(* IEC 61131-3 sources: 2026_Projet_YGO_ExcavatriceDragage/TOOLS/TEST_AUTO_CI/RESULTS/G_CYCLE/reports (part 2) *)

(* ---- FB_CycleSemiAuto_test.st ---- *)
SETUP
VAR
    FB : FB_CycleSemiAuto;
    SampleCount : INT := 0;
    SampleCountTotal : UDINT := 0;
END_VAR
END_SETUP

TEST 'T262-002 AX10B : transfert Both P1 sans coupure M2 puis AX11 P2'
    (* Chargement securise de AX10B : consigne de forcage ecrite par l'operateur (T358). *)
    FB(Enable := TRUE, PowerContactorEngaged := TRUE, Mode := E_Mode.SEMI_AUTO,
       HeartbeatIhmOk := TRUE, M1_SpeedValid := TRUE, M2_SpeedValid := TRUE,
       M1_ContactorsReleased := TRUE, M2_ContactorsReleased := TRUE,
       M1_BrakeApplied := TRUE, M2_BrakeApplied := TRUE,
       M1_MeasuredSpeedMps := 0.0, M2_MeasuredSpeedMps := 0.0,
       JoystickDeflected := FALSE, DeadmanArmed := FALSE,
       CfgCommissioningEnable := TRUE, CfgCtrlAscentMaxStep := 2,
       CfgCtrlAscentDistanceM := 2.0, SampleCount := SampleCount, StepForceTgt := 22);
    ASSERT_TRUE(FB.ForceStepAccepted, 'AX10B forcee immediatement (T358)');
    ASSERT_TRUE(FB.StepForceTgtTaken, 'Consigne vue par le FB : PRG_03 l acquitte (T358)');

    (* Scans d acquittement puis d execution : aucun mouvement au chargement. *)
    FB(StepForceTgt := -1, SampleCount := SampleCount);
    FB(SampleCount := SampleCount);
    ASSERT_FALSE(FB.WinchM1Cmd.RunRequest OR FB.WinchM2Cmd.RunRequest,
                 'Chargement AX10B sans mouvement');

    (* Nouveau geste Y+ : M1 et M2 sont publies simultanement a P1. *)
    FB(StartCycle := FALSE, JoystickDeflected := TRUE, DeadmanArmed := TRUE,
       JoystickPull := TRUE, M2_SpeedStepApplied := 1,
       M1FinalAscentStartReady := TRUE, Benne_CloseReached := TRUE,
       Benne_IsClosed := TRUE, Benne_IsRoughlyClosed := TRUE,
       SampleCount := SampleCount);
    ASSERT_TRUE(FB.CycleStep = E_AutoCycleStep.AX10B_RACCORDEMENT_P1,
                'Scan transfert execute en AX10B');
    ASSERT_TRUE(FB.WinchM1Cmd.RunRequest AND FB.WinchM2Cmd.RunRequest,
                'AX10B publie Both sans trou de commande');
    ASSERT_TRUE((FB.WinchM1Cmd.StepTgt = 1) AND (FB.WinchM2Cmd.StepTgt = 1),
                'AX10B publie M1 P1 et M2 P1');
    ASSERT_TRUE(FB.WinchM1Cmd.ReqAscent AND FB.WinchM2Cmd.ReqAscent,
                'AX10B conserve le sens montee des deux treuils');

    (* Scan suivant : AX11 reprend avec le plafond commun configure P2. *)
    FB(SampleCount := SampleCount);
    ASSERT_TRUE(FB.CycleStep = E_AutoCycleStep.AX11_CTRL_ASCENT,
                'AX11 prend le relais apres transfert P1/P1');
    ASSERT_TRUE((FB.WinchM1Cmd.StepTgt = 2) AND (FB.WinchM2Cmd.StepTgt = 2),
                'AX11 applique le plafond commun P2');
END_TEST

(* ============================================================================
   T345-L2 - AX14->AX15A instantane, neutre obligatoire avant AX15B
   Contrat : TASK_CONTRACT_T345_L2_AX14_AX15A_INSTANTANEE.yaml
   ============================================================================ *)

TEST 'T345-L2-001 : arrivee AX14 neutre, puis nouveau push autorise AX15B'
    FB(Enable := TRUE, PowerContactorEngaged := TRUE, Mode := E_Mode.SEMI_AUTO,
       HeartbeatIhmOk := TRUE, M1_SpeedValid := TRUE, M2_SpeedValid := TRUE,
       M1_ContactorsReleased := TRUE, M2_ContactorsReleased := TRUE,
       M1_BrakeApplied := TRUE, M2_BrakeApplied := TRUE,
       HomedM1 := TRUE, HomedM2 := TRUE, InitPositionOk := TRUE, WinchesAtTopWindow := TRUE,
       Translation_At_Tremie := TRUE, Translation_Busy := FALSE,
       JoystickDeflected := FALSE, DeadmanArmed := TRUE,
       JoystickPush := FALSE, JoystickPull := FALSE, JoystickLeft := FALSE, JoystickRight := FALSE,
       SampleCount := SampleCount, StepForceTgt := 14);
    ASSERT_TRUE(FB.ForceStepAccepted, 'T345-L2-001 : AX14 force');
    FB(StepForceTgt := -1, Translation_At_Tremie := TRUE, Translation_Busy := FALSE,
       JoystickDeflected := FALSE, DeadmanArmed := TRUE, JoystickPush := FALSE,
       SampleCount := SampleCount);
    ADVANCE_TIME(600000000);
    FB(Translation_At_Tremie := TRUE, Translation_Busy := FALSE,
       JoystickDeflected := FALSE, DeadmanArmed := TRUE, JoystickPush := FALSE,
       SampleCount := SampleCount);

    (* Premier scan AX15A au neutre : le latch s'arme, sans transition dans ce meme scan. *)
    FB(Translation_At_Tremie := TRUE, Translation_Busy := FALSE,
       JoystickDeflected := FALSE, DeadmanArmed := TRUE, JoystickPush := FALSE,
       SampleCount := SampleCount);
    ASSERT_TRUE(FB.CycleStep = E_AutoCycleStep.AX15A_DUMP_ARRIVE,
                'T345-L2-001 : AX15A atteint apres confirmation arret');
    ASSERT_FALSE(FB.BucketCmd.ReqOpen OR FB.WinchM1Cmd.RunRequest OR FB.WinchM2Cmd.RunRequest OR FB.TranslationCmd.ReqStart,
                 'T345-L2-001 : aucune commande au scan neutre AX15A');
    ASSERT_EQ(FB.OperatorAction, 'AX15a - Pousser vers le bas pour ouvrir et vider.',
              'T345-L2-001 : guide push publie apres neutre');

    (* Nouveau geste : changement d'etat, puis commande seulement au scan AX15B. *)
    FB(JoystickDeflected := TRUE, DeadmanArmed := TRUE, JoystickPush := TRUE,
       SampleCount := SampleCount);
    ASSERT_TRUE(FB.CycleStep = E_AutoCycleStep.AX15A_DUMP_ARRIVE,
                'T345-L2-001 : transition demandee depuis AX15A');
    ASSERT_FALSE(FB.BucketCmd.ReqOpen, 'T345-L2-001 : aucune ouverture au scan de transition');
    FB(JoystickDeflected := TRUE, DeadmanArmed := TRUE, JoystickPush := TRUE,
       SampleCount := SampleCount);
    ASSERT_TRUE(FB.CycleStep = E_AutoCycleStep.AX15B_DUMP_OPEN,
                'T345-L2-001 : AX15B execute au scan suivant');
    ASSERT_TRUE(FB.BucketCmd.ReqOpen, 'T345-L2-001 : ouverture autorisee apres neutre puis nouveau push');
END_TEST

TEST 'T345-L2-002 : push Y maintenu a l arrivee passe AX15A mais reste bloque avant neutre'
    FB(Enable := TRUE, PowerContactorEngaged := TRUE, Mode := E_Mode.SEMI_AUTO,
       HeartbeatIhmOk := TRUE, M1_SpeedValid := TRUE, M2_SpeedValid := TRUE,
       M1_ContactorsReleased := TRUE, M2_ContactorsReleased := TRUE,
       M1_BrakeApplied := TRUE, M2_BrakeApplied := TRUE,
       HomedM1 := TRUE, HomedM2 := TRUE, InitPositionOk := TRUE, WinchesAtTopWindow := TRUE,
       Translation_At_Tremie := TRUE, Translation_Busy := FALSE,
       JoystickDeflected := TRUE, DeadmanArmed := TRUE,
       JoystickPush := TRUE, JoystickPull := FALSE, JoystickLeft := FALSE, JoystickRight := FALSE,
       SampleCount := SampleCount, StepForceTgt := 14);
    FB(StepForceTgt := -1, Translation_At_Tremie := TRUE, Translation_Busy := FALSE,
       JoystickDeflected := TRUE, DeadmanArmed := TRUE, JoystickPush := TRUE,
       SampleCount := SampleCount);
    ADVANCE_TIME(600000000);
    FB(Translation_At_Tremie := TRUE, Translation_Busy := FALSE,
       JoystickDeflected := TRUE, DeadmanArmed := TRUE, JoystickPush := TRUE,
       SampleCount := SampleCount);
    FB(Translation_At_Tremie := TRUE, Translation_Busy := FALSE,
       JoystickDeflected := TRUE, DeadmanArmed := TRUE, JoystickPush := TRUE,
       SampleCount := SampleCount);
    ASSERT_TRUE(FB.CycleStep = E_AutoCycleStep.AX15A_DUMP_ARRIVE,
                'T345-L2-002 : transition AX14->AX15A sans attendre neutre');
    ASSERT_TRUE(FB.WaitingForOperator, 'T345-L2-002 : relachement operateur attendu');
    ASSERT_EQ(FB.OperatorAction, 'AX15a - Relacher le joystick avant ouverture.',
              'T345-L2-002 : message de relachement explicite');
    ASSERT_FALSE(FB.BucketCmd.ReqOpen OR FB.WinchM1Cmd.RunRequest OR FB.WinchM2Cmd.RunRequest OR FB.TranslationCmd.ReqStart,
                 'T345-L2-002 : Y maintenu ne commande aucun mouvement avant neutre');
    FB(JoystickDeflected := TRUE, DeadmanArmed := TRUE, JoystickPush := TRUE,
       SampleCount := SampleCount);
    ASSERT_TRUE(FB.CycleStep = E_AutoCycleStep.AX15A_DUMP_ARRIVE,
                'T345-L2-002 : AX15A maintenu tant que Y reste pousse');
    ASSERT_FALSE(FB.BucketCmd.ReqOpen, 'T345-L2-002 : ReqOpen reste faux avant neutre');
END_TEST

TEST 'T345-L2-003 : diagonale X plus Y maintenue ne contourne pas le neutre AX15A'
    FB(Enable := TRUE, PowerContactorEngaged := TRUE, Mode := E_Mode.SEMI_AUTO,
       HeartbeatIhmOk := TRUE, M1_SpeedValid := TRUE, M2_SpeedValid := TRUE,
       M1_ContactorsReleased := TRUE, M2_ContactorsReleased := TRUE,
       M1_BrakeApplied := TRUE, M2_BrakeApplied := TRUE,
       HomedM1 := TRUE, HomedM2 := TRUE, InitPositionOk := TRUE, WinchesAtTopWindow := TRUE,
       Translation_At_Tremie := TRUE, Translation_Busy := FALSE,
       JoystickDeflected := TRUE, DeadmanArmed := TRUE,
       JoystickPush := TRUE, JoystickPull := FALSE, JoystickLeft := TRUE, JoystickRight := FALSE,
       SampleCount := SampleCount, StepForceTgt := 14);
    FB(StepForceTgt := -1, Translation_At_Tremie := TRUE, Translation_Busy := FALSE,
       JoystickDeflected := TRUE, DeadmanArmed := TRUE, JoystickPush := TRUE, JoystickLeft := TRUE,
       SampleCount := SampleCount);
    ADVANCE_TIME(600000000);
    FB(Translation_At_Tremie := TRUE, Translation_Busy := FALSE,
       JoystickDeflected := TRUE, DeadmanArmed := TRUE, JoystickPush := TRUE, JoystickLeft := TRUE,
       SampleCount := SampleCount);
    FB(Translation_At_Tremie := TRUE, Translation_Busy := FALSE,
       JoystickDeflected := TRUE, DeadmanArmed := TRUE, JoystickPush := TRUE, JoystickLeft := TRUE,
       SampleCount := SampleCount);
    ASSERT_TRUE(FB.CycleStep = E_AutoCycleStep.AX15A_DUMP_ARRIVE,
                'T345-L2-003 : diagonale n empeche pas l arrivee AX15A');
    ASSERT_FALSE(FB.BucketCmd.ReqOpen OR FB.WinchM1Cmd.RunRequest OR FB.WinchM2Cmd.RunRequest OR FB.TranslationCmd.ReqStart,
                 'T345-L2-003 : diagonale ne produit aucun mouvement avant neutre');
    FB(JoystickDeflected := TRUE, DeadmanArmed := TRUE, JoystickPush := TRUE, JoystickLeft := TRUE,
       SampleCount := SampleCount);
    ASSERT_TRUE(FB.CycleStep = E_AutoCycleStep.AX15A_DUMP_ARRIVE,
                'T345-L2-003 : diagonale maintenue reste bloquee en AX15A');
    ASSERT_FALSE(FB.BucketCmd.ReqOpen, 'T345-L2-003 : ReqOpen reste faux sous diagonale');
END_TEST

TEST 'T345-L2-004 : forcage repete cible 15 efface un latch neutre precedent'
    FB(Enable := TRUE, PowerContactorEngaged := TRUE, Mode := E_Mode.SEMI_AUTO,
       HeartbeatIhmOk := TRUE, M1_SpeedValid := TRUE, M2_SpeedValid := TRUE,
       M1_ContactorsReleased := TRUE, M2_ContactorsReleased := TRUE,
       M1_BrakeApplied := TRUE, M2_BrakeApplied := TRUE,
       HomedM1 := TRUE, HomedM2 := TRUE, InitPositionOk := TRUE, WinchesAtTopWindow := TRUE,
       JoystickDeflected := FALSE, DeadmanArmed := TRUE, JoystickPush := FALSE,
       SampleCount := SampleCount, StepForceTgt := 15);
    FB(StepForceTgt := -1, JoystickDeflected := FALSE, DeadmanArmed := TRUE, JoystickPush := FALSE,
       SampleCount := SampleCount);
    ASSERT_TRUE(FB.CycleStep = E_AutoCycleStep.AX15A_DUMP_ARRIVE,
                'T345-L2-004 : AX15A execute au neutre et latch arme');

    (* Meme cible forcee pendant un push : le reset doit avoir lieu meme sans changement d enum. *)
    FB(StepForceTgt := 15, JoystickDeflected := TRUE, DeadmanArmed := TRUE, JoystickPush := TRUE,
       SampleCount := SampleCount);
    ASSERT_TRUE(FB.ForceStepAccepted, 'T345-L2-004 : forcage repete 15 accepte et neutre en commandes');
    ASSERT_FALSE(FB.BucketCmd.ReqOpen, 'T345-L2-004 : scan de forcage sans ouverture');
    FB(StepForceTgt := -1, JoystickDeflected := TRUE, DeadmanArmed := TRUE, JoystickPush := TRUE,
       SampleCount := SampleCount);
    FB(JoystickDeflected := TRUE, DeadmanArmed := TRUE, JoystickPush := TRUE,
       SampleCount := SampleCount);
    ASSERT_TRUE(FB.CycleStep = E_AutoCycleStep.AX15A_DUMP_ARRIVE,
                'T345-L2-004 : latch perime ne survit pas au forcage repete');
    ASSERT_FALSE(FB.BucketCmd.ReqOpen, 'T345-L2-004 : push deja actif reste bloque sans nouveau neutre');
END_TEST

TEST 'T345-L2-005 : non regression AX2 vers AX3 conserve le geste PushOnly existant'
    FB(Enable := TRUE, PowerContactorEngaged := TRUE, Mode := E_Mode.SEMI_AUTO,
       HeartbeatIhmOk := TRUE, M1_SpeedValid := TRUE, M2_SpeedValid := TRUE,
       M1_ContactorsReleased := TRUE, M2_ContactorsReleased := TRUE,
       M1_BrakeApplied := TRUE, M2_BrakeApplied := TRUE,
       HomedM1 := TRUE, HomedM2 := TRUE, InitPositionOk := TRUE, WinchesAtTopWindow := TRUE,
       Translation_At_P1 := TRUE, Translation_Busy := FALSE,
       JoystickDeflected := TRUE, DeadmanArmed := TRUE,
       JoystickPush := TRUE, JoystickPull := FALSE, JoystickLeft := FALSE, JoystickRight := FALSE,
       SampleCount := SampleCount, StepForceTgt := 2);
    FB(StepForceTgt := -1, Translation_At_P1 := TRUE, Translation_Busy := FALSE,
       JoystickDeflected := TRUE, DeadmanArmed := TRUE, JoystickPush := TRUE,
       JoystickLeft := FALSE, JoystickRight := FALSE, SampleCount := SampleCount);
    ADVANCE_TIME(600000000);
    FB(Translation_At_P1 := TRUE, Translation_Busy := FALSE,
       JoystickDeflected := TRUE, DeadmanArmed := TRUE, JoystickPush := TRUE,
       JoystickLeft := FALSE, JoystickRight := FALSE, SampleCount := SampleCount);
    FB(Translation_At_P1 := TRUE, Translation_Busy := FALSE,
       JoystickDeflected := TRUE, DeadmanArmed := TRUE, JoystickPush := TRUE,
       JoystickLeft := FALSE, JoystickRight := FALSE, SampleCount := SampleCount);
    ASSERT_TRUE(FB.CycleStep = E_AutoCycleStep.AX3_OPEN_BUCKET,
                'T345-L2-005 : AX2->AX3 PushOnly inchange');
    ASSERT_TRUE(FB.BucketCmd.ReqOpen, 'T345-L2-005 : AX3 ouvre comme avant');
END_TEST

TEST 'T262-003 AX10B : timeout M1 borne a 2 s puis repli sans redemarrage implicite'
    (* Preparation AX10B au neutre, comme pour le test nominal (T358). *)
    FB(Enable := TRUE, PowerContactorEngaged := TRUE, Mode := E_Mode.SEMI_AUTO,
       HeartbeatIhmOk := TRUE, M1_SpeedValid := TRUE, M2_SpeedValid := TRUE,
       M1_ContactorsReleased := TRUE, M2_ContactorsReleased := TRUE,
       M1_BrakeApplied := TRUE, M2_BrakeApplied := TRUE,
       M1_MeasuredSpeedMps := 0.0, M2_MeasuredSpeedMps := 0.0,
       JoystickDeflected := FALSE, DeadmanArmed := FALSE,
       CfgCommissioningEnable := TRUE, CfgCtrlAscentMaxStep := 2,
       CfgCtrlAscentDistanceM := 2.0, SampleCount := SampleCount, StepForceTgt := 22);
    ASSERT_TRUE(FB.ForceStepAccepted, 'AX10B forcee pour test timeout (T358)');
    ASSERT_TRUE(FB.StepForceTgtTaken, 'Consigne vue par le FB : PRG_03 l acquitte (T358)');
    FB(StepForceTgt := -1, SampleCount := SampleCount);
    FB(SampleCount := SampleCount);

    (* M1 indisponible : M2 est tenu en P1 pendant la fenetre bornee. *)
    FB(StartCycle := FALSE, JoystickDeflected := TRUE, DeadmanArmed := TRUE,
       JoystickPull := TRUE, M2_SpeedStepApplied := 1,
       M1FinalAscentStartReady := FALSE, Benne_CloseReached := TRUE,
       Benne_IsClosed := TRUE, Benne_IsRoughlyClosed := TRUE,
       SampleCount := SampleCount);
    ASSERT_TRUE(FB.BucketCmd.ReqHoldAscentP1AfterClose,
                'Fenetre AX10B : maintien P1 actif avant timeout');

    ADVANCE_TIME(2100000000);
    FB(SampleCount := SampleCount);
    ASSERT_FALSE(FB.BucketCmd.ReqHoldAscentP1AfterClose,
                 'Timeout : maintien M2 libere');
    ASSERT_FALSE(FB.WinchM1Cmd.RunRequest OR FB.WinchM2Cmd.RunRequest,
                 'Timeout : aucun redemarrage pendant arret de repli');

    ADVANCE_TIME(600000000);
    FB(SampleCount := SampleCount);
    ASSERT_TRUE(FB.CycleStep = E_AutoCycleStep.AX10B_RACCORDEMENT_P1,
                'Repli : AX10B conserve la main pendant la confirmation arret');
    ADVANCE_TIME(600000000);
    FB(SampleCount := SampleCount);
    ASSERT_TRUE(FB.CycleStep = E_AutoCycleStep.AX10B_RACCORDEMENT_P1,
                'Repli : dernier scan AX10B avant reprise');
    FB(SampleCount := SampleCount);
    ASSERT_TRUE(FB.CycleStep = E_AutoCycleStep.AX11_CTRL_ASCENT,
                'Repli : reprise explicite par AX11');
    ASSERT_TRUE(FB.WinchM1Cmd.RunRequest AND FB.WinchM2Cmd.RunRequest,
                'Repli : AX11 reprend les deux treuils ensemble');
END_TEST

TEST 'T331-001 AX15d micro-step benne : tirer ouvre le module, pousser ouvrir, relacher retour AX15B'
    SampleCount := 0;

    (* Chargement securise de l etape de vidage au joystick neutre, machine arretee. *)
    FB(Enable := TRUE, Reset := FALSE, PowerContactorEngaged := TRUE, Mode := E_Mode.SEMI_AUTO,
       HeartbeatIhmOk := TRUE, M1_SpeedValid := TRUE, M2_SpeedValid := TRUE,
       M1_ContactorsReleased := TRUE, M2_ContactorsReleased := TRUE,
       M1_BrakeApplied := TRUE, M2_BrakeApplied := TRUE,
       M1_MeasuredSpeedMps := 0.0, M2_MeasuredSpeedMps := 0.0,
       M1_SpeedStepApplied := 1, M2_SpeedStepApplied := 1,
       JoystickDeflected := FALSE, DeadmanArmed := FALSE,
       JoystickPush := FALSE, JoystickPull := FALSE, JoystickRight := FALSE, JoystickLeft := FALSE,
       StartCycle := FALSE, AbortCycle := FALSE,
       SpeedMismatchThresholdMps := 0.0, SpeedMismatchTimeout := T#0ms,
       WinchSyncError := FALSE, WinchSyncDeltaM := 0.0,
       HomedM1 := TRUE, HomedM2 := TRUE, InitPositionOk := TRUE, WinchesAtTopWindow := TRUE,
       M1_CablePosM := 7.0, M2_CablePosM := 7.0,
       Translation_At_P1 := FALSE, Translation_At_Tremie := TRUE, Translation_At_Maintenance := FALSE,
       Translation_Busy := FALSE, Translation_Done := TRUE,
       Benne_Busy := FALSE, Benne_Done := FALSE, Benne_CloseReached := FALSE,
       Benne_IsOpen := FALSE, Benne_IsClosed := FALSE, Benne_IsRoughlyClosed := FALSE,
       RepositionRequest := FALSE, SkipDrainRequest := FALSE, CfgDrainTime := T#0s,
       CfgCommissioningEnable := TRUE,
       CfgCtrlAscentMaxStep := 1, CfgCtrlAscentDistanceM := 2.0,
       SampleCount := SampleCount);
    FB(StepForceTgt := 16, SampleCount := SampleCount);
    ASSERT_TRUE(FB.ForceStepAccepted, 'Etape de vidage forcee (T331-001)');
    FB(StepForceTgt := -1, SampleCount := SampleCount);
    FB(SampleCount := SampleCount);

    (* Geste nominal maintenu Y- : vidage, treuils neutralises, aucune transition. *)
    FB(StartCycle := FALSE, JoystickDeflected := TRUE, DeadmanArmed := TRUE,
       JoystickPush := TRUE, SampleCount := SampleCount);
    ASSERT_TRUE(FB.CycleStep = E_AutoCycleStep.AX15B_DUMP_OPEN, 'Vidage observe');
    ASSERT_TRUE(FB.BucketCmd.ReqOpen, 'Vidage : ouverture benne commandee');
    ASSERT_FALSE(FB.BucketCmd.ReqClose, 'Vidage : aucune fermeture benne commandee');
    ASSERT_FALSE(FB.WinchM1Cmd.RunRequest OR FB.WinchM2Cmd.RunRequest,
                 'Vidage : les deux treuils restent neutralises');

    (* T383 : tirer ne fait PLUS de saut AX15B -> AX10. Il entre dans le micro-step AX15D. *)
    FB(JoystickPush := FALSE, JoystickPull := TRUE, SampleCount := SampleCount);
    FB(SampleCount := SampleCount);
    ASSERT_TRUE(FB.CycleStep = E_AutoCycleStep.AX15D_DUMP_BUCKET_JOG,
                'T383 : tirer entre dans le micro-step benne AX15D');
    ASSERT_FALSE(FB.CycleStep = E_AutoCycleStep.AX10_CLOSE_BUCKET,
                 'T383 : AUCUN saut vers AX10 (decharge non declaree retiree)');
    ASSERT_FALSE(FB.BucketCmd.ReqOpen, 'AX15D : ouverture neutralisee au tirer');
    ASSERT_TRUE(FB.BucketCmd.ReqClose, 'AX15D : tirer ferme la benne');
    ASSERT_FALSE(FB.WinchM1Cmd.RunRequest OR FB.WinchM2Cmd.RunRequest,
                 'AX15D : les deux treuils restent a 0 (aucun mouvement)');

    (* Module : pousser dans AX15D rouvre la benne, treuils toujours 0. *)
    FB(JoystickPush := TRUE, JoystickPull := FALSE, SampleCount := SampleCount);
    ASSERT_TRUE(FB.CycleStep = E_AutoCycleStep.AX15D_DUMP_BUCKET_JOG,
                'AX15D : on reste dans le micro-step pendant la manipulation');
    ASSERT_TRUE(FB.BucketCmd.ReqOpen, 'AX15D : pousser ouvre la benne');
    ASSERT_FALSE(FB.BucketCmd.ReqClose, 'AX15D : aucune fermeture simultanee');
    ASSERT_FALSE(FB.WinchM1Cmd.RunRequest OR FB.WinchM2Cmd.RunRequest,
                 'AX15D : treuils neutralises pendant le module');

    (* Retour au centre mort : on reprend le vidage (AX15B) sans remontee. *)
    FB(JoystickPush := FALSE, JoystickPull := FALSE, JoystickDeflected := FALSE,
       SampleCount := SampleCount);
    FB(SampleCount := SampleCount);   // AX15D assigne State:=AX15B -> CycleStep au scan suivant
    ASSERT_TRUE(FB.CycleStep = E_AutoCycleStep.AX15B_DUMP_OPEN,
                'AX15D : relachement -> retour au vidage AX15B');
    ASSERT_FALSE(FB.BucketCmd.ReqOpen OR FB.BucketCmd.ReqClose,
                 'AX15D : neutre = les deux demandes benne a zero');
    ASSERT_FALSE(FB.WinchM1Cmd.RunRequest OR FB.WinchM2Cmd.RunRequest,
                 'AX15D : aucun treuil commande au relachement');

    (* Fin de vidage : la benne ouverte amene AX18 sur geste pousse, inchange. *)
    FB(Benne_Done := TRUE, Benne_IsOpen := TRUE, Benne_IsClosed := FALSE,
       Benne_IsRoughlyClosed := FALSE, JoystickDeflected := TRUE, JoystickPush := TRUE,
       SampleCount := SampleCount);
    FB(SampleCount := SampleCount);
    ASSERT_TRUE(FB.CycleStep = E_AutoCycleStep.AX18_DONE_SYNC,
                'Fin de vidage apres module : AX18 inchange');
    ASSERT_FALSE(FB.BucketCmd.ReqOpen, 'Fin de vidage : ouverture relachee');
END_TEST

TEST 'T331-002 AX15b/AX15c non-regression : vidage nominal et repositionnement inchanges'
    SampleCount := 0;

    (* Chargement securise de l etape de vidage au joystick neutre. *)
    FB(Enable := TRUE, Reset := FALSE, PowerContactorEngaged := TRUE, Mode := E_Mode.SEMI_AUTO,
       HeartbeatIhmOk := TRUE, M1_SpeedValid := TRUE, M2_SpeedValid := TRUE,
       M1_ContactorsReleased := TRUE, M2_ContactorsReleased := TRUE,
       M1_BrakeApplied := TRUE, M2_BrakeApplied := TRUE,
       M1_MeasuredSpeedMps := 0.0, M2_MeasuredSpeedMps := 0.0,
       M1_SpeedStepApplied := 1, M2_SpeedStepApplied := 1,
       JoystickDeflected := FALSE, DeadmanArmed := FALSE,
       JoystickPush := FALSE, JoystickPull := FALSE, JoystickRight := FALSE, JoystickLeft := FALSE,
       StartCycle := FALSE, AbortCycle := FALSE,
       SpeedMismatchThresholdMps := 0.0, SpeedMismatchTimeout := T#0ms,
       WinchSyncError := FALSE, WinchSyncDeltaM := 0.0,
       HomedM1 := TRUE, HomedM2 := TRUE, InitPositionOk := TRUE, WinchesAtTopWindow := TRUE,
       M1_CablePosM := 7.0, M2_CablePosM := 7.0,
       Translation_At_P1 := FALSE, Translation_At_Tremie := TRUE, Translation_At_Maintenance := FALSE,
       Translation_Busy := FALSE, Translation_Done := TRUE,
       Benne_Busy := FALSE, Benne_Done := FALSE, Benne_CloseReached := FALSE,
       Benne_IsOpen := FALSE, Benne_IsClosed := FALSE, Benne_IsRoughlyClosed := FALSE,
       RepositionRequest := FALSE, SkipDrainRequest := FALSE, CfgDrainTime := T#0s,
       CfgCommissioningEnable := TRUE,
       CfgCtrlAscentMaxStep := 1, CfgCtrlAscentDistanceM := 2.0,
       SampleCount := SampleCount);
    FB(StepForceTgt := 16, SampleCount := SampleCount);
    ASSERT_TRUE(FB.ForceStepAccepted, 'Etape de vidage forcee (non-regression T358)');
    ASSERT_TRUE(FB.StepForceTgtTaken, 'Consigne vue par le FB : PRG_03 l acquitte (T358)');
    FB(StepForceTgt := -1, SampleCount := SampleCount);

    (* Vidage nominal Y- : ouverture seule, treuils neutralises. *)
    FB(StartCycle := FALSE, JoystickDeflected := TRUE, DeadmanArmed := TRUE,
       JoystickPush := TRUE, SampleCount := SampleCount);
    ASSERT_TRUE(FB.CycleStep = E_AutoCycleStep.AX15B_DUMP_OPEN, 'Vidage nominal inchange');
    ASSERT_TRUE(FB.BucketCmd.ReqOpen, 'Vidage nominal : ouverture commandee');
    ASSERT_FALSE(FB.BucketCmd.ReqClose, 'Vidage nominal : aucune fermeture');
    ASSERT_FALSE(FB.WinchM1Cmd.RunRequest OR FB.WinchM2Cmd.RunRequest,
                 'Vidage nominal : treuils a l arret');

    (* Option IHM maintenue : repositionnement couple en descente, inchange. *)
    FB(RepositionRequest := TRUE, SampleCount := SampleCount);
    FB(SampleCount := SampleCount);
    ASSERT_TRUE(FB.CycleStep = E_AutoCycleStep.AX15C_DUMP_REPOSITION,
                'Repositionnement inchange : AX15c atteint');
    ASSERT_TRUE(FB.WinchM1Cmd.RunRequest AND FB.WinchM2Cmd.RunRequest,
                'Repositionnement : M1 et M2 commandes');
    ASSERT_TRUE(FB.WinchM1Cmd.ReqDescend AND FB.WinchM2Cmd.ReqDescend,
                'Repositionnement : descente couplee conservee');
    ASSERT_FALSE(FB.WinchM1Cmd.ReqAscent OR FB.WinchM2Cmd.ReqAscent,
                 'Repositionnement : aucune montee commandee');
    ASSERT_EQ(FB.WinchM1Cmd.StepTgt, FB.WinchM2Cmd.StepTgt,
              'Repositionnement : meme palier M1/M2');

    (* Relachement de l option : retour au vidage, treuils de nouveau a l arret. *)
    FB(RepositionRequest := FALSE, SampleCount := SampleCount);
    FB(SampleCount := SampleCount);
    ASSERT_TRUE(FB.CycleStep = E_AutoCycleStep.AX15B_DUMP_OPEN,
                'Retour au vidage inchange au relachement de l option');
    ASSERT_FALSE(FB.WinchM1Cmd.RunRequest OR FB.WinchM2Cmd.RunRequest,
                 'Retour vidage : treuils arretes');

    (* Vidage termine : la benne ouverte amene la fin de passe, inchange. *)
    FB(Benne_Done := TRUE, Benne_IsOpen := TRUE, Benne_IsClosed := FALSE,
       Benne_IsRoughlyClosed := FALSE, SampleCount := SampleCount);
    FB(SampleCount := SampleCount);
    ASSERT_TRUE(FB.CycleStep = E_AutoCycleStep.AX18_DONE_SYNC, 'Fin de vidage inchangee');
    ASSERT_FALSE(FB.BucketCmd.ReqOpen, 'Fin de vidage : ouverture relachee');
    ASSERT_EQ(FB.SampleCount, 1, 'Fin de vidage : compteur incremente une seule fois');
END_TEST

TEST 'T331-003 AX15d micro-step : perte du geste, de l homme-mort ou defaut neutralise sans reprise'
    SampleCount := 0;

    (* Chargement securise de l etape de vidage au joystick neutre. *)
    FB(Enable := TRUE, Reset := FALSE, PowerContactorEngaged := TRUE, Mode := E_Mode.SEMI_AUTO,
       HeartbeatIhmOk := TRUE, M1_SpeedValid := TRUE, M2_SpeedValid := TRUE,
       M1_ContactorsReleased := TRUE, M2_ContactorsReleased := TRUE,
       M1_BrakeApplied := TRUE, M2_BrakeApplied := TRUE,
       M1_MeasuredSpeedMps := 0.0, M2_MeasuredSpeedMps := 0.0,
       M1_SpeedStepApplied := 1, M2_SpeedStepApplied := 1,
       JoystickDeflected := FALSE, DeadmanArmed := FALSE,
       JoystickPush := FALSE, JoystickPull := FALSE, JoystickRight := FALSE, JoystickLeft := FALSE,
       StartCycle := FALSE, AbortCycle := FALSE,
       SpeedMismatchThresholdMps := 0.0, SpeedMismatchTimeout := T#0ms,
       WinchSyncError := FALSE, WinchSyncDeltaM := 0.0,
       HomedM1 := TRUE, HomedM2 := TRUE, InitPositionOk := TRUE, WinchesAtTopWindow := TRUE,
       M1_CablePosM := 7.0, M2_CablePosM := 7.0,
       Translation_At_P1 := FALSE, Translation_At_Tremie := TRUE, Translation_At_Maintenance := FALSE,
       Translation_Busy := FALSE, Translation_Done := TRUE,
       Benne_Busy := FALSE, Benne_Done := FALSE, Benne_CloseReached := FALSE,
       Benne_IsOpen := FALSE, Benne_IsClosed := FALSE, Benne_IsRoughlyClosed := FALSE,
       RepositionRequest := FALSE, SkipDrainRequest := FALSE, CfgDrainTime := T#0s,
       CfgCommissioningEnable := TRUE,
       CfgCtrlAscentMaxStep := 1, CfgCtrlAscentDistanceM := 2.0,
       SampleCount := SampleCount);
    FB(StepForceTgt := 16, SampleCount := SampleCount);
    ASSERT_TRUE(FB.ForceStepAccepted, 'Etape de vidage forcee (T331-003)');
    FB(StepForceTgt := -1, SampleCount := SampleCount);
    FB(SampleCount := SampleCount);

    (* Vidage puis tirer maintenu : entre dans le micro-step AX15D, fermeture commandee. *)
    FB(StartCycle := FALSE, JoystickDeflected := TRUE, DeadmanArmed := TRUE,
       JoystickPush := TRUE, SampleCount := SampleCount);
    FB(JoystickPush := FALSE, JoystickPull := TRUE, SampleCount := SampleCount);
    FB(SampleCount := SampleCount);
    ASSERT_TRUE(FB.CycleStep = E_AutoCycleStep.AX15D_DUMP_BUCKET_JOG,
                'Micro-step : entree dans AX15D au tirer');
    ASSERT_TRUE(FB.BucketCmd.ReqClose, 'Micro-step : fermeture benne commandee au tirer');

    (* Relachement du manche : plus aucune demande, retour au vidage AX15B. *)
    FB(JoystickDeflected := FALSE, JoystickPull := FALSE, DeadmanArmed := TRUE,
       SampleCount := SampleCount);
    ASSERT_FALSE(FB.BucketCmd.ReqClose, 'Relachement : fermeture benne neutralisee');
    ASSERT_FALSE(FB.WinchM1Cmd.RunRequest OR FB.WinchM2Cmd.RunRequest,
                 'Relachement : treuils neutralises');
    FB(SampleCount := SampleCount);
    ASSERT_TRUE(FB.CycleStep = E_AutoCycleStep.AX15B_DUMP_OPEN,
                'Relachement : retour a AX15B (reprendre le vidage)');
    ASSERT_FALSE(FB.BucketCmd.ReqClose, 'Relachement : aucune reprise automatique');

    (* Geste repris (tirer) : retour dans le micro-step sous commande maintenue. *)
    FB(JoystickDeflected := TRUE, JoystickPull := TRUE, SampleCount := SampleCount);
    FB(SampleCount := SampleCount);
    ASSERT_TRUE(FB.CycleStep = E_AutoCycleStep.AX15D_DUMP_BUCKET_JOG,
                'Geste repris : retour dans AX15D');
    ASSERT_TRUE(FB.BucketCmd.ReqClose, 'Geste repris : fermeture benne reprise');

    (* Perte de l homme-mort : neutralisation complete, etape conservee. *)
    FB(DeadmanArmed := FALSE, SampleCount := SampleCount);
    ASSERT_FALSE(FB.BucketCmd.ReqClose OR FB.BucketCmd.ReqOpen
                 OR FB.WinchM1Cmd.RunRequest OR FB.WinchM2Cmd.RunRequest,
                 'Homme-mort perdu : plus aucune demande de mouvement');
    FB(SampleCount := SampleCount);
    ASSERT_TRUE(FB.CycleStep = E_AutoCycleStep.AX15D_DUMP_BUCKET_JOG,
                'Homme-mort perdu : etape conservee, aucune reprise automatique');

    (* Defaut pendant le micro-step : repli AX_STAB, sorties neutralisees. *)
    FB(DeadmanArmed := TRUE, HeartbeatIhmOk := FALSE, SampleCount := SampleCount);
    ASSERT_TRUE(FB.CycleStep = E_AutoCycleStep.AX_STAB, 'Defaut : repli AX_STAB');
    ASSERT_FALSE(FB.BucketCmd.ReqClose OR FB.BucketCmd.ReqOpen
                 OR FB.WinchM1Cmd.RunRequest OR FB.WinchM2Cmd.RunRequest,
                 'Defaut : toutes les demandes neutralisees');
    ASSERT_FALSE(FB.Lifecycle.Busy, 'Defaut : cycle non actif');

    (* Acquittement conscient : cause disparue puis Reset. *)
    FB(HeartbeatIhmOk := TRUE, JoystickDeflected := FALSE, JoystickPull := FALSE,
       DeadmanArmed := FALSE, Reset := TRUE, SampleCount := SampleCount);
    FB(Reset := FALSE, SampleCount := SampleCount);
    ASSERT_FALSE(FB.Fault.Latched, 'Acquittement : defaut efface apres cause disparue');
    ASSERT_TRUE(FB.CycleStep = E_AutoCycleStep.AX0_REPOS, 'Acquittement : retour au repos');
END_TEST

TEST 'TC-P03-001 Dynamique Enable : neutralisation initiale, transition Ready au repos, puis coupure'
    (* Scan 0 : Enable=FALSE -> Neutralisation *)
    FB(Enable := FALSE, Reset := FALSE, PowerContactorEngaged := TRUE, Mode := E_Mode.SEMI_AUTO,
       DeadmanArmed := FALSE, JoystickDeflected := FALSE, JoystickPush := FALSE, M1_SpeedValid := TRUE, M2_SpeedValid := TRUE, M1_ContactorsReleased := TRUE, M2_ContactorsReleased := TRUE, M1_BrakeApplied := TRUE, M2_BrakeApplied := TRUE, M1_SpeedStepApplied := 4, M2_SpeedStepApplied := 4, HeartbeatIhmOk := TRUE,
       StartCycle := FALSE, SampleCount := SampleCount);
    ASSERT_FALSE(FB.Ready, 'Enable=FALSE -> Ready=FALSE (neutralise)');
    ASSERT_FALSE(FB.Lifecycle.Busy, 'Enable=FALSE -> Lifecycle.Busy=FALSE');

    ADVANCE_TIME(10000000);

    (* Scan 1 : Enable=TRUE -> Prete en service *)
    FB(Enable := TRUE, Reset := FALSE, PowerContactorEngaged := TRUE, Mode := E_Mode.SEMI_AUTO,
       DeadmanArmed := FALSE, JoystickDeflected := FALSE, JoystickPush := FALSE, M1_SpeedValid := TRUE, M2_SpeedValid := TRUE, M1_ContactorsReleased := TRUE, M2_ContactorsReleased := TRUE, M1_BrakeApplied := TRUE, M2_BrakeApplied := TRUE, M1_SpeedStepApplied := 4, M2_SpeedStepApplied := 4, HeartbeatIhmOk := TRUE,
       StartCycle := FALSE, SampleCount := SampleCount);
    ASSERT_TRUE(FB.Ready, 'Enable=TRUE -> Ready=TRUE (nominal)');
    ASSERT_FALSE(FB.Lifecycle.Busy, 'Au repos -> Pas de cycle actif');

    ADVANCE_TIME(10000000);

    (* Scan 2 : Enable=FALSE -> Re-neutralisation *)
    FB(Enable := FALSE, Reset := FALSE, PowerContactorEngaged := TRUE, Mode := E_Mode.SEMI_AUTO,
       DeadmanArmed := FALSE, JoystickDeflected := FALSE, JoystickPush := FALSE, M1_SpeedValid := TRUE, M2_SpeedValid := TRUE, M1_ContactorsReleased := TRUE, M2_ContactorsReleased := TRUE, M1_BrakeApplied := TRUE, M2_BrakeApplied := TRUE, M1_SpeedStepApplied := 4, M2_SpeedStepApplied := 4, HeartbeatIhmOk := TRUE,
       StartCycle := FALSE, SampleCount := SampleCount);
    ASSERT_FALSE(FB.Ready, 'Coupure -> Ready retombe a FALSE');
END_TEST

TEST 'TC-P04-027 T258 : ForÃ§age prepare sans action et reprise sur Start au neutre'
    (* T358 : consigne unique ecrite par l'operateur — AUCUNE condition de contexte,
       aucune confirmation. Le joystick est volontairement DEFLECHI pour prouver que la
       garde « joystick au neutre » a bien disparu, et l'homme-mort reste absent pour
       verifier que le forcage lui-meme ne cree AUCUN mouvement. *)
    FB(Enable := TRUE, PowerContactorEngaged := TRUE, Mode := E_Mode.SEMI_AUTO,
       HeartbeatIhmOk := TRUE, M1_SpeedValid := TRUE, M2_SpeedValid := TRUE,
       M1_ContactorsReleased := TRUE, M2_ContactorsReleased := TRUE,
       M1_BrakeApplied := TRUE, M2_BrakeApplied := TRUE,
       JoystickDeflected := TRUE, DeadmanArmed := FALSE,
       CfgCommissioningEnable := TRUE, SampleCount := SampleCount, StepForceTgt := 4);
    ASSERT_TRUE(FB.ForceStepAccepted, 'Saut accepte joystick deflechi, sans aucune condition (T358)');
    ASSERT_TRUE(FB.StepForceTgtTaken, 'Consigne vue par le FB : PRG_03 l acquitte (T358)');
    ASSERT_FALSE(FB.WinchM1Cmd.RunRequest OR FB.WinchM2Cmd.RunRequest, 'Aucune action au scan du forcage');
    FB(StepForceTgt := -1, SampleCount := SampleCount);
    ASSERT_TRUE(FB.CycleStep = E_AutoCycleStep.AX4_DESCEND_DIVING, 'AX4 chargee au scan suivant (T358)');
    ASSERT_FALSE(FB.WinchM1Cmd.RunRequest OR FB.WinchM2Cmd.RunRequest, 'Le forcage ne cree aucun mouvement');
    FB(StartCycle := FALSE, DeadmanArmed := TRUE, JoystickDeflected := TRUE,
       JoystickPull := TRUE, JoystickPush := FALSE, SampleCount := SampleCount);
    ASSERT_FALSE(FB.WinchM1Cmd.RunRequest OR FB.WinchM2Cmd.RunRequest, 'Y+ ne commande pas la descente AX4');
    FB(JoystickPull := FALSE, JoystickPush := TRUE, SampleCount := SampleCount);
    ASSERT_TRUE(FB.WinchM1Cmd.RunRequest AND FB.WinchM2Cmd.RunRequest, 'Y- commande les deux voies AX4');
END_TEST

TEST 'TC-P04-028 T258 : ForÃ§age AX_STAB refuse et reste neutre'
    (* T358 : AX_STAB (19) etait explicitement REFUSE par l ancienne garde « <> 19 »
       alors que c est une valeur d enum valide : elle est desormais forcable. *)
    FB(Enable := TRUE, PowerContactorEngaged := TRUE, Mode := E_Mode.SEMI_AUTO,
       HeartbeatIhmOk := TRUE, M1_SpeedValid := TRUE, M2_SpeedValid := TRUE,
       M1_ContactorsReleased := TRUE, M2_ContactorsReleased := TRUE,
       M1_BrakeApplied := TRUE, M2_BrakeApplied := TRUE,
       JoystickDeflected := FALSE, CfgCommissioningEnable := TRUE, SampleCount := SampleCount,
       StepForceTgt := 19);
    ASSERT_TRUE(FB.ForceStepAccepted, 'AX_STAB desormais forcable : 19 est dans la plage enum (T358)');
    ASSERT_TRUE(FB.StepForceTgtTaken, 'Consigne vue par le FB : PRG_03 l acquitte (T358)');
    ASSERT_FALSE(FB.ForceStepRejected, 'Aucun rejet d une valeur d enum valide (T358)');
    ASSERT_FALSE(FB.WinchM1Cmd.RunRequest OR FB.WinchM2Cmd.RunRequest, 'Sorties neutres au scan du forcage');
    FB(StepForceTgt := -1, SampleCount := SampleCount);
    ASSERT_TRUE(FB.CycleStep = E_AutoCycleStep.AX_STAB, 'AX_STAB chargee au scan suivant (T358)');
END_TEST

TEST 'TC-P04-029 T258 : Inhibition ne masque pas le desynchronisme'
    FB(Enable := TRUE, PowerContactorEngaged := TRUE, Mode := E_Mode.SEMI_AUTO,
       HeartbeatIhmOk := TRUE, M1_SpeedValid := TRUE, M2_SpeedValid := TRUE,
       M1_ContactorsReleased := TRUE, M2_ContactorsReleased := TRUE,
       M1_BrakeApplied := TRUE, M2_BrakeApplied := TRUE,
       CfgCommissioningEnable := TRUE, CfgCycleChecksInhibit := FALSE,
       StartCycle := TRUE, SampleCount := SampleCount);
    FB(StartCycle := FALSE, CfgCycleChecksInhibit := TRUE, SampleCount := SampleCount);
    ASSERT_TRUE(FB.CycleChecksInhibited, 'Mode essai actif');
    FB(CfgCycleChecksInhibit := TRUE, WinchSyncError := TRUE, SampleCount := SampleCount);
    ASSERT_TRUE(FB.CycleChecksInhibited, 'Mode essai reste actif pendant injection safety');
    ASSERT_TRUE(FB.Fault.Error, 'Synchronisme reste bloquant');
    ASSERT_TRUE(FB.CycleStep = E_AutoCycleStep.AX_STAB, 'Repli AX_STAB maintenu');
END_TEST

TEST 'TC-P04-030 T258 : Un forçage refuse invalide une preparation precedente'
    (* T358 : la SEULE validation restante est la plage de l enum. Hors plage = rejet,
       etape inchangee, consigne acquittee (donc jamais rejouee en boucle). *)
    FB(Enable := TRUE, PowerContactorEngaged := TRUE, Mode := E_Mode.SEMI_AUTO,
       HeartbeatIhmOk := TRUE, M1_SpeedValid := TRUE, M2_SpeedValid := TRUE,
       M1_ContactorsReleased := TRUE, M2_ContactorsReleased := TRUE,
       M1_BrakeApplied := TRUE, M2_BrakeApplied := TRUE,
       JoystickDeflected := FALSE, CfgCommissioningEnable := TRUE,
       StartCycle := FALSE, SampleCount := SampleCount, StepForceTgt := 40);
    ASSERT_TRUE(FB.ForceStepRejected, 'Cible hors plage refusee (T358)');
    ASSERT_FALSE(FB.ForceStepAccepted, 'Aucune consigne appliquee hors plage');
    ASSERT_TRUE(FB.ForceStepResult <> '', 'Motif de rejet publie (T358)');
    ASSERT_TRUE(FB.StepForceTgtTaken, 'Consigne vue par le FB : PRG_03 l acquitte (T358)');
    ASSERT_FALSE(FB.CycleStep = E_AutoCycleStep.AX4_DESCEND_DIVING, 'Aucune etape chargee apres rejet');
    ASSERT_FALSE(FB.WinchM1Cmd.RunRequest OR FB.WinchM2Cmd.RunRequest, 'Start ne peut executer aucune cible');
    (* La consigne acquittee, le scan suivant repart de la sentinelle : aucun rejeu. *)
    FB(StepForceTgt := -1, SampleCount := SampleCount);
    ASSERT_FALSE(FB.ForceStepRejected, 'Impulsion de rejet d un seul scan (T358)');
    FB(StartCycle := FALSE, DeadmanArmed := TRUE, JoystickDeflected := TRUE,
       JoystickPush := TRUE, SampleCount := SampleCount);
    ASSERT_FALSE(FB.WinchM1Cmd.RunRequest OR FB.WinchM2Cmd.RunRequest, 'Nouveau geste Y- sans cible reste neutre');
    ASSERT_FALSE(FB.TranslationCmd.ReqStart OR FB.BucketCmd.ReqOpen OR FB.BucketCmd.ReqClose OR FB.BucketCmd.ReqKoboldMeasureEnable,
                 'Tous les autres actionneurs restent neutres apres rejet');
END_TEST

TEST 'TC-P04-031 T258 : Apply et Start simultanes restent en preparation neutre'
    (* T358 : AX18_DONE_SYNC (18) etait explicitement REFUSE par l ancienne garde
       « <> 18 » alors que c est une valeur d enum valide : elle est desormais forcable. *)
    FB(Enable := TRUE, PowerContactorEngaged := TRUE, Mode := E_Mode.SEMI_AUTO,
       HeartbeatIhmOk := TRUE, M1_SpeedValid := TRUE, M2_SpeedValid := TRUE,
       M1_ContactorsReleased := TRUE, M2_ContactorsReleased := TRUE,
       M1_BrakeApplied := TRUE, M2_BrakeApplied := TRUE,
       JoystickDeflected := FALSE, CfgCommissioningEnable := TRUE,
       StartCycle := FALSE, SampleCount := SampleCount, StepForceTgt := 18);
    ASSERT_TRUE(FB.ForceStepAccepted, 'AX18 forcee : 18 est dans la plage enum (T358)');
    ASSERT_TRUE(FB.StepForceTgtTaken, 'Consigne vue par le FB : PRG_03 l acquitte (T358)');
    ASSERT_FALSE(FB.ForceStepRejected, 'Aucun rejet d une valeur d enum valide (T358)');
    ASSERT_FALSE(FB.WinchM1Cmd.RunRequest OR FB.WinchM2Cmd.RunRequest, 'Aucune commande au scan du forcage');
    FB(StepForceTgt := -1, StartCycle := FALSE, SampleCount := SampleCount);
    ASSERT_TRUE(FB.CycleStep = E_AutoCycleStep.AX18_DONE_SYNC, 'AX18 chargee au scan suivant (T358)');
    ASSERT_FALSE(FB.TranslationCmd.ReqStart OR FB.BucketCmd.ReqOpen OR FB.BucketCmd.ReqClose OR FB.BucketCmd.ReqKoboldMeasureEnable,
                 'Aucun autre actionneur commande par le forcage (T358)');
END_TEST

TEST 'TC-P04-032 T258 : Reset simultane annule le forçage'
    (* T358 : une consigne ecrite sur le MEME scan qu un Reset est effacee par le Reset
       (l abandon et l acquittement precedent le bloc de forcage dans l ordre intra-scan) :
       aucun saut d etape ne peut survivre a un acquittement. *)
    FB(Enable := TRUE, PowerContactorEngaged := TRUE, Mode := E_Mode.SEMI_AUTO,
       HeartbeatIhmOk := TRUE, M1_SpeedValid := TRUE, M2_SpeedValid := TRUE,
       M1_ContactorsReleased := TRUE, M2_ContactorsReleased := TRUE,
       M1_BrakeApplied := TRUE, M2_BrakeApplied := TRUE,
       JoystickDeflected := FALSE, CfgCommissioningEnable := TRUE, Reset := TRUE,
       SampleCount := SampleCount, StepForceTgt := 4);
    ASSERT_TRUE(FB.StepForceTgtTaken, 'Consigne vue par le FB : PRG_03 l acquitte (T358)');
    ASSERT_FALSE(FB.ForceStepAccepted, 'Aucun forcage applique : le Reset du meme scan neutralise la consigne');
    ASSERT_FALSE(FB.CycleStep = E_AutoCycleStep.AX4_DESCEND_DIVING, 'AX4 non chargee apres Reset + consigne');
    FB(StepForceTgt := -1, Reset := FALSE, SampleCount := SampleCount);
    ASSERT_FALSE(FB.CycleStep = E_AutoCycleStep.AX4_DESCEND_DIVING, 'Aucun saut differe au scan suivant (T358)');
END_TEST

TEST 'TC-P04-033 T258 : Forcage semi-auto independant du bit commissioning'
    (* T358 : une consigne ecrite alors que le CYCLE est inactif (hors SEMI_AUTO) est
       ECARTEE — acquittee et motif publie. Elle n est JAMAIS honoree plus tard, a la
       reactivation du cycle : ce serait un saut d etape sans geste nouveau. *)
    FB(Enable := FALSE, PowerContactorEngaged := TRUE, Mode := E_Mode.MAINT_N1,
       HeartbeatIhmOk := TRUE, M1_SpeedValid := TRUE, M2_SpeedValid := TRUE,
       M1_ContactorsReleased := TRUE, M2_ContactorsReleased := TRUE,
       M1_BrakeApplied := TRUE, M2_BrakeApplied := TRUE,
       JoystickDeflected := FALSE, CfgCommissioningEnable := TRUE, SampleCount := SampleCount,
       StepForceTgt := 4);
    ASSERT_TRUE(FB.ForceStepRejected, 'Consigne ecartee : cycle inactif (T358)');
    ASSERT_TRUE(FB.StepForceTgtTaken, 'Consigne vue par le FB : PRG_03 l acquitte (T358)');
    ASSERT_TRUE(FB.ForceStepResult <> '', 'Motif d ecart publie (T358)');
    FB(Enable := TRUE, Mode := E_Mode.SEMI_AUTO, StepForceTgt := -1, SampleCount := SampleCount);
    ASSERT_FALSE(FB.CycleStep = E_AutoCycleStep.AX4_DESCEND_DIVING, 'Aucun saut differe a la reactivation (T358)');
    (* Le forcage reste possible des que le cycle est actif : meme cible, meme scan. *)
    FB(StepForceTgt := 4, SampleCount := SampleCount);
    ASSERT_TRUE(FB.ForceStepAccepted, 'Forcage effectif une fois le cycle actif (T358)');
END_TEST

TEST 'TC-P04-001 : Relachement manche (JoystickDeflected=FALSE) stoppe les commandes sans perdre l etape'
    SampleCount := 5;
    // Initialisation et dÃƒÆ’Ã†â€™Ãƒâ€šÃ‚Â©marrage cycle
    FB(Enable := TRUE, PowerContactorEngaged := TRUE, Mode := E_Mode.SEMI_AUTO,
       DeadmanArmed := TRUE, JoystickDeflected := TRUE, JoystickPush := TRUE, M1_SpeedValid := TRUE, M2_SpeedValid := TRUE, M1_ContactorsReleased := TRUE, M2_ContactorsReleased := TRUE, M1_BrakeApplied := TRUE, M2_BrakeApplied := TRUE, M1_SpeedStepApplied := 4, M2_SpeedStepApplied := 4, HeartbeatIhmOk := TRUE,
       StartCycle := TRUE, SampleCount := SampleCount);

    // Simuler le relÃƒÆ’Ã†â€™Ãƒâ€šÃ‚Â¢chement du manche au centre (JoystickDeflected -> FALSE)
    FB(Enable := TRUE, PowerContactorEngaged := TRUE, Mode := E_Mode.SEMI_AUTO,
       DeadmanArmed := TRUE, JoystickDeflected := FALSE, JoystickPush := FALSE, M1_SpeedValid := TRUE, M2_SpeedValid := TRUE, M1_ContactorsReleased := TRUE, M2_ContactorsReleased := TRUE, M1_BrakeApplied := TRUE, M2_BrakeApplied := TRUE, M1_SpeedStepApplied := 4, M2_SpeedStepApplied := 4, HeartbeatIhmOk := TRUE,
       StartCycle := FALSE, SampleCount := SampleCount);

    ASSERT_FALSE(FB.WinchM1Cmd.RunRequest, 'M1 coupe sur retour neutre manche');
    ASSERT_FALSE(FB.WinchM2Cmd.RunRequest, 'M2 coupe sur retour neutre manche');
    ASSERT_FALSE(FB.TranslationCmd.ReqStart, 'Translation coupee');
    ASSERT_TRUE(FB.CycleStep = E_AutoCycleStep.AX0_REPOS OR FB.CycleStep = E_AutoCycleStep.AX1_INIT, 'Etape conservee');
END_TEST

TEST 'TC-P04-002 : Le cycle produit des demandes et passe a AX1_INIT sur Start'
    SampleCount := 0;
    // Scan 1 : front montant StartCycle -> transition State vers AX1_INIT
    FB(Enable := TRUE, PowerContactorEngaged := TRUE, Mode := E_Mode.SEMI_AUTO,
       DeadmanArmed := TRUE, JoystickDeflected := TRUE, JoystickPush := TRUE, M1_SpeedValid := TRUE, M2_SpeedValid := TRUE, M1_ContactorsReleased := TRUE, M2_ContactorsReleased := TRUE, M1_BrakeApplied := TRUE, M2_BrakeApplied := TRUE, M1_SpeedStepApplied := 4, M2_SpeedStepApplied := 4, HeartbeatIhmOk := TRUE,
       StartCycle := TRUE, SampleCount := SampleCount);

    // Scan 2 : exÃƒÆ’Ã†â€™Ãƒâ€šÃ‚Â©cution de l'ÃƒÆ’Ã†â€™Ãƒâ€šÃ‚Â©tape AX1_INIT -> Lifecycle.Busy=TRUE
    FB(Enable := TRUE, PowerContactorEngaged := TRUE, Mode := E_Mode.SEMI_AUTO,
       DeadmanArmed := TRUE, JoystickDeflected := TRUE, JoystickPush := TRUE, M1_SpeedValid := TRUE, M2_SpeedValid := TRUE, M1_ContactorsReleased := TRUE, M2_ContactorsReleased := TRUE, M1_BrakeApplied := TRUE, M2_BrakeApplied := TRUE, M1_SpeedStepApplied := 4, M2_SpeedStepApplied := 4, HeartbeatIhmOk := TRUE,
       StartCycle := FALSE, SampleCount := SampleCount);

    ASSERT_TRUE(FB.Lifecycle.Busy, 'Cycle actif (Lifecycle.Busy=TRUE)');
    ASSERT_FALSE(FB.Fault.Error, 'Pas d erreur au lancement');
    ASSERT_TRUE(FB.CycleStep = E_AutoCycleStep.AX1_INIT, 'Transition vers AX1_INIT');
END_TEST

TEST 'TC-P04-003 : Defaut de synchronisation treuils bascule le cycle en AX_STAB et fige l etape'
    SampleCount := 0;
    // Scan 1 : DÃƒÆ’Ã†â€™Ãƒâ€šÃ‚Â©marrage
    FB(Enable := TRUE, PowerContactorEngaged := TRUE, Mode := E_Mode.SEMI_AUTO,
       DeadmanArmed := TRUE, JoystickDeflected := TRUE, JoystickPush := TRUE, M1_SpeedValid := TRUE, M2_SpeedValid := TRUE, M1_ContactorsReleased := TRUE, M2_ContactorsReleased := TRUE, M1_BrakeApplied := TRUE, M2_BrakeApplied := TRUE, M1_SpeedStepApplied := 4, M2_SpeedStepApplied := 4, HeartbeatIhmOk := TRUE,
       StartCycle := TRUE, SampleCount := SampleCount);

    // Scan 2 : ÃƒÆ’Ã†â€™ÃƒÂ¢Ã¢â€šÂ¬Ã‚Â°tablissement ÃƒÆ’Ã†â€™Ãƒâ€šÃ‚Â  AX1_INIT
    FB(Enable := TRUE, PowerContactorEngaged := TRUE, Mode := E_Mode.SEMI_AUTO,
       DeadmanArmed := TRUE, JoystickDeflected := TRUE, JoystickPush := TRUE, M1_SpeedValid := TRUE, M2_SpeedValid := TRUE, M1_ContactorsReleased := TRUE, M2_ContactorsReleased := TRUE, M1_BrakeApplied := TRUE, M2_BrakeApplied := TRUE, M1_SpeedStepApplied := 4, M2_SpeedStepApplied := 4, HeartbeatIhmOk := TRUE,
       StartCycle := FALSE, SampleCount := SampleCount);

    // Scan 3 : Injection dÃƒÆ’Ã†â€™Ãƒâ€šÃ‚Â©synchronisme bloquant WinchSyncError
    FB(Enable := TRUE, PowerContactorEngaged := TRUE, Mode := E_Mode.SEMI_AUTO,
       DeadmanArmed := TRUE, JoystickDeflected := TRUE, JoystickPush := TRUE, M1_SpeedValid := TRUE, M2_SpeedValid := TRUE, M1_ContactorsReleased := TRUE, M2_ContactorsReleased := TRUE, M1_BrakeApplied := TRUE, M2_BrakeApplied := TRUE, M1_SpeedStepApplied := 4, M2_SpeedStepApplied := 4, HeartbeatIhmOk := TRUE,
       StartCycle := FALSE, WinchSyncError := TRUE, SampleCount := SampleCount);

    ASSERT_TRUE(FB.CycleStep = E_AutoCycleStep.AX_STAB, 'Bascule en AX_STAB');
    ASSERT_TRUE(FB.Fault.Error, 'Drapeau Fault.Error actif');
    ASSERT_FALSE(FB.WinchM1Cmd.RunRequest, 'Commandes treuils neutralisees');
END_TEST

TEST 'TC-P04-004 : Reprise apres AX_STAB necessite Cause disparue + Reset + StartCycle'
    SampleCount := 0;
    // Scan 1 : Demarrage
    FB(Enable := TRUE, PowerContactorEngaged := TRUE, Mode := E_Mode.SEMI_AUTO,
       DeadmanArmed := TRUE, JoystickDeflected := TRUE, JoystickPush := TRUE, M1_SpeedValid := TRUE, M2_SpeedValid := TRUE, M1_ContactorsReleased := TRUE, M2_ContactorsReleased := TRUE, M1_BrakeApplied := TRUE, M2_BrakeApplied := TRUE, M1_SpeedStepApplied := 4, M2_SpeedStepApplied := 4, HeartbeatIhmOk := TRUE,
       StartCycle := TRUE, SampleCount := SampleCount);
    // Scan 2 : Etablissement a AX1_INIT
    FB(Enable := TRUE, PowerContactorEngaged := TRUE, Mode := E_Mode.SEMI_AUTO,
       DeadmanArmed := TRUE, JoystickDeflected := TRUE, JoystickPush := TRUE, M1_SpeedValid := TRUE, M2_SpeedValid := TRUE, M1_ContactorsReleased := TRUE, M2_ContactorsReleased := TRUE, M1_BrakeApplied := TRUE, M2_BrakeApplied := TRUE, M1_SpeedStepApplied := 4, M2_SpeedStepApplied := 4, HeartbeatIhmOk := TRUE,
       StartCycle := FALSE, SampleCount := SampleCount);
    // Scan 3 : Injection defaut de synchronisme -> Bascule en AX_STAB
    FB(Enable := TRUE, PowerContactorEngaged := TRUE, Mode := E_Mode.SEMI_AUTO,
       DeadmanArmed := TRUE, JoystickDeflected := TRUE, JoystickPush := TRUE, M1_SpeedValid := TRUE, M2_SpeedValid := TRUE, M1_ContactorsReleased := TRUE, M2_ContactorsReleased := TRUE, M1_BrakeApplied := TRUE, M2_BrakeApplied := TRUE, M1_SpeedStepApplied := 4, M2_SpeedStepApplied := 4, HeartbeatIhmOk := TRUE,
       StartCycle := FALSE, WinchSyncError := TRUE, SampleCount := SampleCount);
    ASSERT_TRUE(FB.CycleStep = E_AutoCycleStep.AX_STAB, 'Bascule en AX_STAB');

    // 1. Cause disparue mais pas de Reset
    FB(Enable := TRUE, PowerContactorEngaged := TRUE, Mode := E_Mode.SEMI_AUTO,
       DeadmanArmed := TRUE, JoystickDeflected := TRUE, JoystickPush := TRUE, M1_SpeedValid := TRUE, M2_SpeedValid := TRUE, M1_ContactorsReleased := TRUE, M2_ContactorsReleased := TRUE, M1_BrakeApplied := TRUE, M2_BrakeApplied := TRUE, M1_SpeedStepApplied := 4, M2_SpeedStepApplied := 4, HeartbeatIhmOk := TRUE,
       WinchSyncError := FALSE, Reset := FALSE, StartCycle := FALSE, SampleCount := SampleCount);
    ASSERT_TRUE(FB.CycleStep = E_AutoCycleStep.AX_STAB, 'Reste en AX_STAB sans Reset');

    // 2. Front Reset (acquittement) -> retourne a AX0_REPOS
    FB(Enable := TRUE, PowerContactorEngaged := TRUE, Mode := E_Mode.SEMI_AUTO,
       DeadmanArmed := TRUE, JoystickDeflected := TRUE, JoystickPush := TRUE, M1_SpeedValid := TRUE, M2_SpeedValid := TRUE, M1_ContactorsReleased := TRUE, M2_ContactorsReleased := TRUE, M1_BrakeApplied := TRUE, M2_BrakeApplied := TRUE, M1_SpeedStepApplied := 4, M2_SpeedStepApplied := 4, HeartbeatIhmOk := TRUE,
       WinchSyncError := FALSE, Reset := TRUE, StartCycle := FALSE, SampleCount := SampleCount);
    ASSERT_TRUE(FB.CycleStep = E_AutoCycleStep.AX0_REPOS, 'Sortie de AX_STAB vers X0 sur Reset');

    // 3. Demande de redemarrage explicite StartCycle (Scan 1: front montant, Scan 2: execution)
    FB(Enable := TRUE, PowerContactorEngaged := TRUE, Mode := E_Mode.SEMI_AUTO,
       DeadmanArmed := TRUE, JoystickDeflected := TRUE, JoystickPush := TRUE, M1_SpeedValid := TRUE, M2_SpeedValid := TRUE, M1_ContactorsReleased := TRUE, M2_ContactorsReleased := TRUE, M1_BrakeApplied := TRUE, M2_BrakeApplied := TRUE, M1_SpeedStepApplied := 4, M2_SpeedStepApplied := 4, HeartbeatIhmOk := TRUE,
       WinchSyncError := FALSE, Reset := FALSE, StartCycle := TRUE, SampleCount := SampleCount);
    FB(Enable := TRUE, PowerContactorEngaged := TRUE, Mode := E_Mode.SEMI_AUTO,
       DeadmanArmed := TRUE, JoystickDeflected := TRUE, JoystickPush := TRUE, M1_SpeedValid := TRUE, M2_SpeedValid := TRUE, M1_ContactorsReleased := TRUE, M2_ContactorsReleased := TRUE, M1_BrakeApplied := TRUE, M2_BrakeApplied := TRUE, M1_SpeedStepApplied := 4, M2_SpeedStepApplied := 4, HeartbeatIhmOk := TRUE,
       WinchSyncError := FALSE, Reset := FALSE, StartCycle := FALSE, SampleCount := SampleCount);
    ASSERT_TRUE(FB.CycleStep = E_AutoCycleStep.AX1_INIT, 'Redemarrage reussi vers AX1_INIT');
END_TEST

TEST 'TC-P04-012 : Compteur de prelevements SampleCount RETAIN incremente sur AX18_DONE_SYNC'
    SampleCount := 10;
    FB(Enable := TRUE, PowerContactorEngaged := TRUE, Mode := E_Mode.SEMI_AUTO,
       SampleCount := SampleCount);
    ASSERT_EQ(FB.SampleCount, 10, 'Compteur SampleCount inaltere hors fin de cycle');
END_TEST

TEST 'TC-P04-013 : Bascule Semi-Auto vers Maintenance preserve l etape et neutralise les demandes sans redemarrage auto'
    SampleCount := 0;
    // 1. Lancement du cycle jusqu'ÃƒÆ’Ã†â€™Ãƒâ€šÃ‚Â  AX1_INIT
    FB(Enable := TRUE, PowerContactorEngaged := TRUE, Mode := E_Mode.SEMI_AUTO,
       DeadmanArmed := TRUE, JoystickDeflected := TRUE, JoystickPush := TRUE, M1_SpeedValid := TRUE, M2_SpeedValid := TRUE, M1_ContactorsReleased := TRUE, M2_ContactorsReleased := TRUE, M1_BrakeApplied := TRUE, M2_BrakeApplied := TRUE, M1_SpeedStepApplied := 4, M2_SpeedStepApplied := 4, HeartbeatIhmOk := TRUE,
       StartCycle := TRUE, SampleCount := SampleCount);
    FB(Enable := TRUE, PowerContactorEngaged := TRUE, Mode := E_Mode.SEMI_AUTO,
       DeadmanArmed := TRUE, JoystickDeflected := TRUE, JoystickPush := TRUE, M1_SpeedValid := TRUE, M2_SpeedValid := TRUE, M1_ContactorsReleased := TRUE, M2_ContactorsReleased := TRUE, M1_BrakeApplied := TRUE, M2_BrakeApplied := TRUE, M1_SpeedStepApplied := 4, M2_SpeedStepApplied := 4, HeartbeatIhmOk := TRUE,
       StartCycle := FALSE, SampleCount := SampleCount);
    ASSERT_TRUE(FB.CycleStep = E_AutoCycleStep.AX1_INIT, 'Etape AX1_INIT active');

    // 2. Bascule en mode MAINTENANCE (Enable := FALSE)
    FB(Enable := FALSE, PowerContactorEngaged := TRUE, Mode := E_Mode.MAINT_N1,
       DeadmanArmed := TRUE, JoystickDeflected := TRUE, JoystickPush := TRUE, M1_SpeedValid := TRUE, M2_SpeedValid := TRUE, M1_ContactorsReleased := TRUE, M2_ContactorsReleased := TRUE, M1_BrakeApplied := TRUE, M2_BrakeApplied := TRUE, M1_SpeedStepApplied := 4, M2_SpeedStepApplied := 4, HeartbeatIhmOk := TRUE,
       StartCycle := FALSE, SampleCount := SampleCount);
    ASSERT_FALSE(FB.Ready, 'Ready retombe hors Semi-Auto');
    ASSERT_FALSE(FB.Lifecycle.Busy, 'Busy=FALSE en Maintenance');
    ASSERT_FALSE(FB.WinchM1Cmd.RunRequest, 'Demandes M1 neutralisees');
    ASSERT_TRUE(FB.CycleStep = E_AutoCycleStep.AX1_INIT, 'Etape AX1_INIT preservee en memoire');

    // 3. Retour en mode SEMI_AUTO (Enable := TRUE) avec manche deflechi : PAS de mouvement spontane
    FB(Enable := TRUE, PowerContactorEngaged := TRUE, Mode := E_Mode.SEMI_AUTO,
       DeadmanArmed := TRUE, JoystickDeflected := TRUE, JoystickPush := TRUE, M1_SpeedValid := TRUE, M2_SpeedValid := TRUE, M1_ContactorsReleased := TRUE, M2_ContactorsReleased := TRUE, M1_BrakeApplied := TRUE, M2_BrakeApplied := TRUE, M1_SpeedStepApplied := 4, M2_SpeedStepApplied := 4, HeartbeatIhmOk := TRUE,
       StartCycle := FALSE, SampleCount := SampleCount);
    ASSERT_TRUE(FB.CycleStep = E_AutoCycleStep.AX1_INIT, 'Toujours a AX1_INIT');
END_TEST

TEST 'TC-P04-020 : Homme-mort relache en cours de plongee X4 -> commandes neutralisees, etape maintenue, PAS de redemarrage auto (T169-A S3)'
    SampleCount := 0;
    // === Progression vers AX4_DESCEND_DIVING (pattern chaine : un call pose State, le suivant observe CycleStep) ===
    (* Call 1 : front StartCycle -> X0->X1 *)
    FB(Enable := TRUE, Reset := FALSE, PowerContactorEngaged := TRUE, Mode := E_Mode.SEMI_AUTO,
       DeadmanArmed := TRUE, JoystickDeflected := TRUE, JoystickPush := TRUE, M1_SpeedValid := TRUE, M2_SpeedValid := TRUE, M1_ContactorsReleased := TRUE, M2_ContactorsReleased := TRUE, M1_BrakeApplied := TRUE, M2_BrakeApplied := TRUE, M1_SpeedStepApplied := 4, M2_SpeedStepApplied := 4, HeartbeatIhmOk := TRUE,
       StartCycle := TRUE, SelTarget := 3, SetDepthM := -10.0,
       LimitLegalDepthM := -10.5, CableLimitM1AscentM := 7.0,
       SpeedMismatchThresholdMps := 0.0, SpeedMismatchTimeout := T#0ms,
       HomedM1 := TRUE, HomedM2 := TRUE, InitPositionOk := TRUE, WinchesAtTopWindow := TRUE, HomingRequest := FALSE,
       M1_CablePosM := 7.0, M2_CablePosM := 7.0, M1_MeasuredSpeedMps := 0.0, M2_MeasuredSpeedMps := 0.0,
WinchSyncError := FALSE, WinchSyncDeltaM := 0.0,
       Translation_At_P1 := FALSE, Translation_At_Tremie := FALSE, Translation_At_Maintenance := FALSE,
       Translation_Busy := FALSE, Translation_Done := FALSE,
       Benne_Busy := FALSE, Benne_Done := FALSE, Benne_IsOpen := FALSE, Benne_IsClosed := TRUE, Benne_IsRoughlyClosed := TRUE,
       SampleCount := SampleCount);
    (* Call 2 : observe X1, deja home -> X2 *)
    FB(Enable := TRUE, Reset := FALSE, PowerContactorEngaged := TRUE, Mode := E_Mode.SEMI_AUTO,
       DeadmanArmed := TRUE, JoystickDeflected := TRUE, JoystickPush := TRUE, M1_SpeedValid := TRUE, M2_SpeedValid := TRUE, M1_ContactorsReleased := TRUE, M2_ContactorsReleased := TRUE, M1_BrakeApplied := TRUE, M2_BrakeApplied := TRUE, M1_SpeedStepApplied := 4, M2_SpeedStepApplied := 4, HeartbeatIhmOk := TRUE,
       StartCycle := FALSE, SelTarget := 3, SetDepthM := -10.0,
       LimitLegalDepthM := -10.5, CableLimitM1AscentM := 7.0,
       SpeedMismatchThresholdMps := 0.0, SpeedMismatchTimeout := T#0ms,
       HomedM1 := TRUE, HomedM2 := TRUE, InitPositionOk := TRUE, WinchesAtTopWindow := TRUE, HomingRequest := FALSE,
       M1_CablePosM := 7.0, M2_CablePosM := 7.0, M1_MeasuredSpeedMps := 0.0, M2_MeasuredSpeedMps := 0.0,
WinchSyncError := FALSE, WinchSyncDeltaM := 0.0,
       Translation_At_P1 := FALSE, Translation_At_Tremie := FALSE, Translation_At_Maintenance := FALSE,
       Translation_Busy := FALSE, Translation_Done := FALSE,
       Benne_Busy := FALSE, Benne_Done := FALSE, Benne_IsOpen := FALSE, Benne_IsClosed := TRUE, Benne_IsRoughlyClosed := TRUE,
       SampleCount := SampleCount);
    (* Call 3 : observe X2, cible P1 atteinte -> X3 *)
    FB(Enable := TRUE, Reset := FALSE, PowerContactorEngaged := TRUE, Mode := E_Mode.SEMI_AUTO,
       DeadmanArmed := TRUE, JoystickDeflected := TRUE, JoystickPush := TRUE, M1_SpeedValid := TRUE, M2_SpeedValid := TRUE, M1_ContactorsReleased := TRUE, M2_ContactorsReleased := TRUE, M1_BrakeApplied := TRUE, M2_BrakeApplied := TRUE, M1_SpeedStepApplied := 4, M2_SpeedStepApplied := 4, HeartbeatIhmOk := TRUE,
       StartCycle := FALSE, SelTarget := 3, SetDepthM := -10.0,
       LimitLegalDepthM := -10.5, CableLimitM1AscentM := 7.0,
       SpeedMismatchThresholdMps := 0.0, SpeedMismatchTimeout := T#0ms,
       HomedM1 := TRUE, HomedM2 := TRUE, InitPositionOk := TRUE, WinchesAtTopWindow := TRUE, HomingRequest := FALSE,
       M1_CablePosM := 7.0, M2_CablePosM := 7.0, M1_MeasuredSpeedMps := 0.0, M2_MeasuredSpeedMps := 0.0,
WinchSyncError := FALSE, WinchSyncDeltaM := 0.0,
       Translation_At_P1 := TRUE, Translation_At_Tremie := FALSE, Translation_At_Maintenance := FALSE,
       Translation_Busy := FALSE, Translation_Done := TRUE,
       Benne_Busy := FALSE, Benne_Done := FALSE, Benne_IsOpen := FALSE, Benne_IsClosed := TRUE, Benne_IsRoughlyClosed := TRUE,
       SampleCount := SampleCount);
    (* Call 4 : observe X3, benne ouverte -> X4 *)
    FB(Enable := TRUE, Reset := FALSE, PowerContactorEngaged := TRUE, Mode := E_Mode.SEMI_AUTO,
       DeadmanArmed := TRUE, JoystickDeflected := TRUE, JoystickPush := TRUE, M1_SpeedValid := TRUE, M2_SpeedValid := TRUE, M1_ContactorsReleased := TRUE, M2_ContactorsReleased := TRUE, M1_BrakeApplied := TRUE, M2_BrakeApplied := TRUE, M1_SpeedStepApplied := 4, M2_SpeedStepApplied := 4, HeartbeatIhmOk := TRUE,
       StartCycle := FALSE, SelTarget := 3, SetDepthM := -10.0,
       LimitLegalDepthM := -10.5, CableLimitM1AscentM := 7.0,
       SpeedMismatchThresholdMps := 0.0, SpeedMismatchTimeout := T#0ms,
       HomedM1 := TRUE, HomedM2 := TRUE, InitPositionOk := TRUE, WinchesAtTopWindow := TRUE, HomingRequest := FALSE,
       M1_CablePosM := 7.0, M2_CablePosM := 7.0, M1_MeasuredSpeedMps := 0.0, M2_MeasuredSpeedMps := 0.0,
WinchSyncError := FALSE, WinchSyncDeltaM := 0.0,
       Translation_At_P1 := TRUE, Translation_At_Tremie := FALSE, Translation_At_Maintenance := FALSE,
       Translation_Busy := FALSE, Translation_Done := TRUE,
       Benne_Busy := FALSE, Benne_Done := FALSE, Benne_IsOpen := TRUE, Benne_IsClosed := FALSE, Benne_IsRoughlyClosed := FALSE,
       SampleCount := SampleCount);
    (* Call 5 : observe AX4_DESCEND_DIVING, plongee sans contact fond *)
    FB(Enable := TRUE, Reset := FALSE, PowerContactorEngaged := TRUE, Mode := E_Mode.SEMI_AUTO,
       DeadmanArmed := TRUE, JoystickDeflected := TRUE, JoystickPush := TRUE, M1_SpeedValid := TRUE, M2_SpeedValid := TRUE, M1_ContactorsReleased := TRUE, M2_ContactorsReleased := TRUE, M1_BrakeApplied := TRUE, M2_BrakeApplied := TRUE, M1_SpeedStepApplied := 4, M2_SpeedStepApplied := 4, HeartbeatIhmOk := TRUE,
       StartCycle := FALSE, SelTarget := 3, SetDepthM := -10.0,
       LimitLegalDepthM := -10.5, CableLimitM1AscentM := 7.0,
       SpeedMismatchThresholdMps := 0.0, SpeedMismatchTimeout := T#0ms,
       HomedM1 := TRUE, HomedM2 := TRUE, InitPositionOk := TRUE, WinchesAtTopWindow := TRUE, HomingRequest := FALSE,
       M1_CablePosM := 5.0, M2_CablePosM := 5.0, M1_MeasuredSpeedMps := 0.0, M2_MeasuredSpeedMps := 0.0,
WinchSyncError := FALSE, WinchSyncDeltaM := 0.0,
       Translation_At_P1 := TRUE, Translation_At_Tremie := FALSE, Translation_At_Maintenance := FALSE,
       Translation_Busy := FALSE, Translation_Done := TRUE,
       Benne_Busy := FALSE, Benne_Done := FALSE, Benne_IsOpen := TRUE, Benne_IsClosed := FALSE, Benne_IsRoughlyClosed := FALSE,
       SampleCount := SampleCount);
    ADVANCE_TIME(300000000);
    FB(SampleCount := SampleCount);
    FB(SampleCount := SampleCount);
    ASSERT_TRUE(FB.CycleStep = E_AutoCycleStep.AX4_DESCEND_DIVING, 'Etabli en AX4_DESCEND_DIVING');
    ASSERT_TRUE(FB.WinchM1Cmd.RunRequest, 'Descente M1 commandee avant relache');
    ASSERT_FALSE(FB.BucketCmd.ReqKoboldMeasureEnable, 'Kobold PAS enclenche en AX4 - enclenche seulement des AX5');
    ASSERT_TRUE(FB.RequestActive, 'RequestActive=TRUE en X4 (plongee active, T186)');

    (* Call 6 : relache homme-mort / manche au centre pendant la plongee -> neutralisation, etape maintenue *)
    FB(Enable := TRUE, Reset := FALSE, PowerContactorEngaged := TRUE, Mode := E_Mode.SEMI_AUTO,
       DeadmanArmed := FALSE, JoystickDeflected := FALSE, JoystickPush := FALSE, M1_SpeedValid := TRUE, M2_SpeedValid := TRUE, M1_ContactorsReleased := TRUE, M2_ContactorsReleased := TRUE, M1_BrakeApplied := TRUE, M2_BrakeApplied := TRUE, M1_SpeedStepApplied := 4, M2_SpeedStepApplied := 4, HeartbeatIhmOk := TRUE,
       StartCycle := FALSE, SelTarget := 3, SetDepthM := -10.0,
       LimitLegalDepthM := -10.5, CableLimitM1AscentM := 7.0,
       SpeedMismatchThresholdMps := 0.0, SpeedMismatchTimeout := T#0ms,
       HomedM1 := TRUE, HomedM2 := TRUE, InitPositionOk := TRUE, WinchesAtTopWindow := TRUE, HomingRequest := FALSE,
       M1_CablePosM := 5.0, M2_CablePosM := 5.0, M1_MeasuredSpeedMps := 0.0, M2_MeasuredSpeedMps := 0.0,
WinchSyncError := FALSE, WinchSyncDeltaM := 0.0,
       Translation_At_P1 := TRUE, Translation_At_Tremie := FALSE, Translation_At_Maintenance := FALSE,
       Translation_Busy := FALSE, Translation_Done := TRUE,
       Benne_Busy := FALSE, Benne_Done := FALSE, Benne_IsOpen := TRUE, Benne_IsClosed := FALSE, Benne_IsRoughlyClosed := FALSE,
       SampleCount := SampleCount);
    ASSERT_FALSE(FB.WinchM1Cmd.RunRequest, 'Descente M1 neutralisee au relache');
    ASSERT_FALSE(FB.WinchM2Cmd.RunRequest, 'Descente M2 neutralisee au relache');
    ASSERT_FALSE(FB.BucketCmd.ReqKoboldMeasureEnable, 'Contacteur Kobold neutralise');
    ASSERT_TRUE(FB.CycleStep = E_AutoCycleStep.AX4_DESCEND_DIVING, 'Etape X4 maintenue (pas de retour X0)');
    ASSERT_FALSE(FB.RequestActive, 'Aucune demande active');

    (* Call 7 : maintient du relache 5 s -> PAS de redemarrage auto, etape figee *)
    ADVANCE_TIME(5000000000);
    FB(Enable := TRUE, Reset := FALSE, PowerContactorEngaged := TRUE, Mode := E_Mode.SEMI_AUTO,
       DeadmanArmed := FALSE, JoystickDeflected := FALSE, JoystickPush := FALSE, M1_SpeedValid := TRUE, M2_SpeedValid := TRUE, M1_ContactorsReleased := TRUE, M2_ContactorsReleased := TRUE, M1_BrakeApplied := TRUE, M2_BrakeApplied := TRUE, M1_SpeedStepApplied := 4, M2_SpeedStepApplied := 4, HeartbeatIhmOk := TRUE,
       StartCycle := FALSE, SelTarget := 3, SetDepthM := -10.0,
       LimitLegalDepthM := -10.5, CableLimitM1AscentM := 7.0,
       SpeedMismatchThresholdMps := 0.0, SpeedMismatchTimeout := T#0ms,
       HomedM1 := TRUE, HomedM2 := TRUE, InitPositionOk := TRUE, WinchesAtTopWindow := TRUE, HomingRequest := FALSE,
       M1_CablePosM := 5.0, M2_CablePosM := 5.0, M1_MeasuredSpeedMps := 0.0, M2_MeasuredSpeedMps := 0.0,
WinchSyncError := FALSE, WinchSyncDeltaM := 0.0,
       Translation_At_P1 := TRUE, Translation_At_Tremie := FALSE, Translation_At_Maintenance := FALSE,
       Translation_Busy := FALSE, Translation_Done := TRUE,
       Benne_Busy := FALSE, Benne_Done := FALSE, Benne_IsOpen := TRUE, Benne_IsClosed := FALSE, Benne_IsRoughlyClosed := FALSE,
       SampleCount := SampleCount);
    ASSERT_TRUE(FB.CycleStep = E_AutoCycleStep.AX4_DESCEND_DIVING, 'Etape X4 figee apres 5 s de relache');
    ASSERT_FALSE(FB.WinchM1Cmd.RunRequest, 'Aucun redemarrage auto M1');
    ASSERT_FALSE(FB.Fault.Error, 'Pas de defaut (le relache homme-mort n est pas un defaut)');

    (* T358 : la reprise consciente apres bascule de mode est CONSERVEE — elle ne passe
       plus par le chemin du forçage, et le scenario « forçage refuse pendant l attente »
       n existe plus : la consigne 19 (AX_STAB) est desormais ACCEPTEE (test T358 dedie).
       Ce bloc verifie donc la reprise consciente SANS aucune consigne de forçage. *)
    FB(Enable := FALSE, Mode := E_Mode.MAINT_N1, JoystickDeflected := FALSE,
       DeadmanArmed := FALSE, JoystickPush := FALSE, CfgCommissioningEnable := TRUE,
       SampleCount := SampleCount);
    FB(Enable := TRUE, Mode := E_Mode.SEMI_AUTO, JoystickDeflected := FALSE,
       DeadmanArmed := FALSE, JoystickPush := FALSE, SampleCount := SampleCount);
    ASSERT_TRUE(FB.CycleStep = E_AutoCycleStep.AX4_DESCEND_DIVING,
                'Etape X4 memorisee : attente de reprise consciente');
    ASSERT_FALSE(FB.WinchM1Cmd.RunRequest OR FB.WinchM2Cmd.RunRequest,
                 'Retour en SEMI_AUTO sans geste : aucune remise en mouvement');
    FB(DeadmanArmed := FALSE, JoystickDeflected := FALSE, JoystickPush := FALSE,
       StartCycle := TRUE, SampleCount := SampleCount);
    ASSERT_FALSE(FB.WinchM1Cmd.RunRequest OR FB.WinchM2Cmd.RunRequest,
                 'Scan Start de reprise reste neutre');

    (* Call 8 : nouveau geste apres Start -> reprise a X4 SANS repartir de X0 *)
    FB(Enable := TRUE, Reset := FALSE, PowerContactorEngaged := TRUE, Mode := E_Mode.SEMI_AUTO,
       DeadmanArmed := TRUE, JoystickDeflected := TRUE, JoystickPush := TRUE, M1_SpeedValid := TRUE, M2_SpeedValid := TRUE, M1_ContactorsReleased := TRUE, M2_ContactorsReleased := TRUE, M1_BrakeApplied := TRUE, M2_BrakeApplied := TRUE, M1_SpeedStepApplied := 4, M2_SpeedStepApplied := 4, HeartbeatIhmOk := TRUE,
       StartCycle := FALSE, SelTarget := 3, SetDepthM := -10.0,
       LimitLegalDepthM := -10.5, CableLimitM1AscentM := 7.0,
       SpeedMismatchThresholdMps := 0.0, SpeedMismatchTimeout := T#0ms,
       HomedM1 := TRUE, HomedM2 := TRUE, InitPositionOk := TRUE, WinchesAtTopWindow := TRUE, HomingRequest := FALSE,
       M1_CablePosM := 5.0, M2_CablePosM := 5.0, M1_MeasuredSpeedMps := 0.0, M2_MeasuredSpeedMps := 0.0,
WinchSyncError := FALSE, WinchSyncDeltaM := 0.0,
       Translation_At_P1 := TRUE, Translation_At_Tremie := FALSE, Translation_At_Maintenance := FALSE,
       Translation_Busy := FALSE, Translation_Done := TRUE,
       Benne_Busy := FALSE, Benne_Done := FALSE, Benne_IsOpen := TRUE, Benne_IsClosed := FALSE, Benne_IsRoughlyClosed := FALSE,
       SampleCount := SampleCount);
    ASSERT_TRUE(FB.CycleStep = E_AutoCycleStep.AX4_DESCEND_DIVING, 'Reprise a X4 (pas de redemarrage depuis X0)');
    ASSERT_TRUE(FB.WinchM1Cmd.RunRequest, 'Descente M1 commandee apres re-armement');
END_TEST

TEST 'TC-P04-021 : Fond jamais atteint -> maintien AX4 car tempo max etape desactivee'
    SampleCount := 0;
    (* === Progression vers AX4_DESCEND_DIVING (KoboldImmersed reste FALSE = sonde hors eau) === *)
    (* Call 1 : front StartCycle -> X0->X1 *)
    FB(Enable := TRUE, Reset := FALSE, PowerContactorEngaged := TRUE, Mode := E_Mode.SEMI_AUTO,
       DeadmanArmed := TRUE, JoystickDeflected := TRUE, JoystickPush := TRUE, M1_SpeedValid := TRUE, M2_SpeedValid := TRUE, M1_ContactorsReleased := TRUE, M2_ContactorsReleased := TRUE, M1_BrakeApplied := TRUE, M2_BrakeApplied := TRUE, M1_SpeedStepApplied := 4, M2_SpeedStepApplied := 4, HeartbeatIhmOk := TRUE,
       StartCycle := TRUE, SelTarget := 3, SetDepthM := -10.0,
       LimitLegalDepthM := -10.5, CableLimitM1AscentM := 7.0, DiveStartMinM := 4.0,
       SpeedMismatchThresholdMps := 0.0, SpeedMismatchTimeout := T#0ms,
       HomedM1 := TRUE, HomedM2 := TRUE, InitPositionOk := TRUE, WinchesAtTopWindow := TRUE, HomingRequest := FALSE,
       M1_CablePosM := 7.0, M2_CablePosM := 7.0, M1_MeasuredSpeedMps := 0.0, M2_MeasuredSpeedMps := 0.0,
WinchSyncError := FALSE, WinchSyncDeltaM := 0.0,
       Translation_At_P1 := FALSE, Translation_At_Tremie := FALSE, Translation_At_Maintenance := FALSE,
       Translation_Busy := FALSE, Translation_Done := FALSE,
       Benne_Busy := FALSE, Benne_Done := FALSE, Benne_IsOpen := FALSE, Benne_IsClosed := TRUE, Benne_IsRoughlyClosed := TRUE,
       SampleCount := SampleCount);
    (* Call 2 : observe X1, deja home -> X2 *)
    FB(Enable := TRUE, Reset := FALSE, PowerContactorEngaged := TRUE, Mode := E_Mode.SEMI_AUTO,
       DeadmanArmed := TRUE, JoystickDeflected := TRUE, JoystickPush := TRUE, M1_SpeedValid := TRUE, M2_SpeedValid := TRUE, M1_ContactorsReleased := TRUE, M2_ContactorsReleased := TRUE, M1_BrakeApplied := TRUE, M2_BrakeApplied := TRUE, M1_SpeedStepApplied := 4, M2_SpeedStepApplied := 4, HeartbeatIhmOk := TRUE,
       StartCycle := FALSE, SelTarget := 3, SetDepthM := -10.0,
       LimitLegalDepthM := -10.5, CableLimitM1AscentM := 7.0, DiveStartMinM := 4.0,
       SpeedMismatchThresholdMps := 0.0, SpeedMismatchTimeout := T#0ms,
       HomedM1 := TRUE, HomedM2 := TRUE, InitPositionOk := TRUE, WinchesAtTopWindow := TRUE, HomingRequest := FALSE,
       M1_CablePosM := 7.0, M2_CablePosM := 7.0, M1_MeasuredSpeedMps := 0.0, M2_MeasuredSpeedMps := 0.0,
WinchSyncError := FALSE, WinchSyncDeltaM := 0.0,
       Translation_At_P1 := FALSE, Translation_At_Tremie := FALSE, Translation_At_Maintenance := FALSE,
       Translation_Busy := FALSE, Translation_Done := FALSE,
       Benne_Busy := FALSE, Benne_Done := FALSE, Benne_IsOpen := FALSE, Benne_IsClosed := TRUE, Benne_IsRoughlyClosed := TRUE,
       SampleCount := SampleCount);
    (* Call 3 : observe X2, cible P1 atteinte -> X3 *)
    FB(Enable := TRUE, Reset := FALSE, PowerContactorEngaged := TRUE, Mode := E_Mode.SEMI_AUTO,
       DeadmanArmed := TRUE, JoystickDeflected := TRUE, JoystickPush := TRUE, M1_SpeedValid := TRUE, M2_SpeedValid := TRUE, M1_ContactorsReleased := TRUE, M2_ContactorsReleased := TRUE, M1_BrakeApplied := TRUE, M2_BrakeApplied := TRUE, M1_SpeedStepApplied := 4, M2_SpeedStepApplied := 4, HeartbeatIhmOk := TRUE,
       StartCycle := FALSE, SelTarget := 3, SetDepthM := -10.0,
       LimitLegalDepthM := -10.5, CableLimitM1AscentM := 7.0, DiveStartMinM := 4.0,
       SpeedMismatchThresholdMps := 0.0, SpeedMismatchTimeout := T#0ms,
       HomedM1 := TRUE, HomedM2 := TRUE, InitPositionOk := TRUE, WinchesAtTopWindow := TRUE, HomingRequest := FALSE,
       M1_CablePosM := 7.0, M2_CablePosM := 7.0, M1_MeasuredSpeedMps := 0.0, M2_MeasuredSpeedMps := 0.0,
WinchSyncError := FALSE, WinchSyncDeltaM := 0.0,
       Translation_At_P1 := TRUE, Translation_At_Tremie := FALSE, Translation_At_Maintenance := FALSE,
       Translation_Busy := FALSE, Translation_Done := TRUE,
       Benne_Busy := FALSE, Benne_Done := FALSE, Benne_IsOpen := FALSE, Benne_IsClosed := TRUE, Benne_IsRoughlyClosed := TRUE,
       SampleCount := SampleCount);
    (* Call 4 : observe X3, benne ouverte -> X4 *)
    FB(Enable := TRUE, Reset := FALSE, PowerContactorEngaged := TRUE, Mode := E_Mode.SEMI_AUTO,
       DeadmanArmed := TRUE, JoystickDeflected := TRUE, JoystickPush := TRUE, M1_SpeedValid := TRUE, M2_SpeedValid := TRUE, M1_ContactorsReleased := TRUE, M2_ContactorsReleased := TRUE, M1_BrakeApplied := TRUE, M2_BrakeApplied := TRUE, M1_SpeedStepApplied := 4, M2_SpeedStepApplied := 4, HeartbeatIhmOk := TRUE,
       StartCycle := FALSE, SelTarget := 3, SetDepthM := -10.0,
       LimitLegalDepthM := -10.5, CableLimitM1AscentM := 7.0, DiveStartMinM := 4.0,
       SpeedMismatchThresholdMps := 0.0, SpeedMismatchTimeout := T#0ms,
       HomedM1 := TRUE, HomedM2 := TRUE, InitPositionOk := TRUE, WinchesAtTopWindow := TRUE, HomingRequest := FALSE,
       M1_CablePosM := 5.0, M2_CablePosM := 5.0, M1_MeasuredSpeedMps := 0.0, M2_MeasuredSpeedMps := 0.0,
WinchSyncError := FALSE, WinchSyncDeltaM := 0.0,
       Translation_At_P1 := TRUE, Translation_At_Tremie := FALSE, Translation_At_Maintenance := FALSE,
       Translation_Busy := FALSE, Translation_Done := TRUE,
       Benne_Busy := FALSE, Benne_Done := FALSE, Benne_IsOpen := TRUE, Benne_IsClosed := FALSE, Benne_IsRoughlyClosed := FALSE,
       SampleCount := SampleCount);
    (* Call 5 : observe AX4_DESCEND_DIVING, plongee sans contact fond (Kobold = FALSE) *)
    FB(Enable := TRUE, Reset := FALSE, PowerContactorEngaged := TRUE, Mode := E_Mode.SEMI_AUTO,
       DeadmanArmed := TRUE, JoystickDeflected := TRUE, JoystickPush := TRUE, M1_SpeedValid := TRUE, M2_SpeedValid := TRUE, M1_ContactorsReleased := TRUE, M2_ContactorsReleased := TRUE, M1_BrakeApplied := TRUE, M2_BrakeApplied := TRUE, M1_SpeedStepApplied := 4, M2_SpeedStepApplied := 4, HeartbeatIhmOk := TRUE,
       StartCycle := FALSE, SelTarget := 3, SetDepthM := -10.0,
       LimitLegalDepthM := -10.5, CableLimitM1AscentM := 7.0, DiveStartMinM := 4.0,
       SpeedMismatchThresholdMps := 0.0, SpeedMismatchTimeout := T#0ms,
       HomedM1 := TRUE, HomedM2 := TRUE, InitPositionOk := TRUE, WinchesAtTopWindow := TRUE, HomingRequest := FALSE,
       M1_CablePosM := 5.0, M2_CablePosM := 5.0, M1_MeasuredSpeedMps := 0.0, M2_MeasuredSpeedMps := 0.0,
WinchSyncError := FALSE, WinchSyncDeltaM := 0.0,
       Translation_At_P1 := TRUE, Translation_At_Tremie := FALSE, Translation_At_Maintenance := FALSE,
       Translation_Busy := FALSE, Translation_Done := TRUE,
       Benne_Busy := FALSE, Benne_Done := FALSE, Benne_IsOpen := TRUE, Benne_IsClosed := FALSE, Benne_IsRoughlyClosed := FALSE,
       SampleCount := SampleCount);
    ADVANCE_TIME(300000000);
    FB(SampleCount := SampleCount);
    FB(SampleCount := SampleCount);
    ASSERT_TRUE(FB.CycleStep = E_AutoCycleStep.AX4_DESCEND_DIVING, 'Etabli en AX4_DESCEND_DIVING');

    (* Call 5bis : 1 scan de stabilisation en X4 -> StepMaxTimer armee (StepMaxPrevState = X4)
       apres le rearmement au changement d'etape. Sans ce scan, la tempo est encore a 0 et
       l'ADVANCE_TIME qui suit ne serait pas compte (IN passe FALSE->TRUE au scan d'avance). *)
    FB(Enable := TRUE, Reset := FALSE, PowerContactorEngaged := TRUE, Mode := E_Mode.SEMI_AUTO,
       DeadmanArmed := TRUE, JoystickDeflected := TRUE, JoystickPush := TRUE, M1_SpeedValid := TRUE, M2_SpeedValid := TRUE, M1_ContactorsReleased := TRUE, M2_ContactorsReleased := TRUE, M1_BrakeApplied := TRUE, M2_BrakeApplied := TRUE, M1_SpeedStepApplied := 4, M2_SpeedStepApplied := 4, HeartbeatIhmOk := TRUE,
       StartCycle := FALSE, SelTarget := 3, SetDepthM := -10.0,
       LimitLegalDepthM := -10.5, CableLimitM1AscentM := 7.0, DiveStartMinM := 4.0,
       SpeedMismatchThresholdMps := 0.0, SpeedMismatchTimeout := T#0ms,
       HomedM1 := TRUE, HomedM2 := TRUE, InitPositionOk := TRUE, WinchesAtTopWindow := TRUE, HomingRequest := FALSE,
       M1_CablePosM := 5.0, M2_CablePosM := 5.0, M1_MeasuredSpeedMps := 0.0, M2_MeasuredSpeedMps := 0.0,
WinchSyncError := FALSE, WinchSyncDeltaM := 0.0,
       Translation_At_P1 := TRUE, Translation_At_Tremie := FALSE, Translation_At_Maintenance := FALSE,
       Translation_Busy := FALSE, Translation_Done := TRUE,
       Benne_Busy := FALSE, Benne_Done := FALSE, Benne_IsOpen := TRUE, Benne_IsClosed := FALSE, Benne_IsRoughlyClosed := FALSE,
       SampleCount := SampleCount);

    (* Call 6 : fond toujours pas atteint -> avance de 61 s (> StepMaxTimeout 60 s) -> timeout etape *)
    ADVANCE_TIME(61000000000);
    FB(Enable := TRUE, Reset := FALSE, PowerContactorEngaged := TRUE, Mode := E_Mode.SEMI_AUTO,
       DeadmanArmed := TRUE, JoystickDeflected := TRUE, JoystickPush := TRUE, M1_SpeedValid := TRUE, M2_SpeedValid := TRUE, M1_ContactorsReleased := TRUE, M2_ContactorsReleased := TRUE, M1_BrakeApplied := TRUE, M2_BrakeApplied := TRUE, M1_SpeedStepApplied := 4, M2_SpeedStepApplied := 4, HeartbeatIhmOk := TRUE,
       StartCycle := FALSE, SelTarget := 3, SetDepthM := -10.0,
       LimitLegalDepthM := -10.5, CableLimitM1AscentM := 7.0, DiveStartMinM := 4.0,
       SpeedMismatchThresholdMps := 0.0, SpeedMismatchTimeout := T#0ms,
       HomedM1 := TRUE, HomedM2 := TRUE, InitPositionOk := TRUE, WinchesAtTopWindow := TRUE, HomingRequest := FALSE,
       M1_CablePosM := 5.0, M2_CablePosM := 5.0, M1_MeasuredSpeedMps := 0.0, M2_MeasuredSpeedMps := 0.0,
WinchSyncError := FALSE, WinchSyncDeltaM := 0.0,
       Translation_At_P1 := TRUE, Translation_At_Tremie := FALSE, Translation_At_Maintenance := FALSE,
       Translation_Busy := FALSE, Translation_Done := TRUE,
       Benne_Busy := FALSE, Benne_Done := FALSE, Benne_IsOpen := TRUE, Benne_IsClosed := FALSE, Benne_IsRoughlyClosed := FALSE,
       SampleCount := SampleCount);
    ASSERT_TRUE(FB.CycleStep = E_AutoCycleStep.AX4_DESCEND_DIVING, 'Tempo max desactivee : AX4 maintenue');
    ASSERT_FALSE(FB.Fault.Error, 'Aucun defaut temporel quand StepMaxTimer est desactive');
    ASSERT_TRUE(FB.WinchM1Cmd.RunRequest, 'Commande M1 maintenue');
    ASSERT_TRUE(FB.WinchM2Cmd.RunRequest, 'Commande M2 maintenue');
    ASSERT_TRUE(FB.RequestActive, 'Demande de plongee active');
    ASSERT_FALSE(FB.Fault.Latched, 'Aucun defaut latche');
    ASSERT_FALSE(FB.BucketCmd.ReqKoboldMeasureEnable, 'Kobold reste coupe en AX4');

END_TEST

TEST 'TC-P04-023 : StepMaxTimer NON cumulatif - 2 etapes de 40 s (total 80 s > 60 s) sans AX_STAB'
    SampleCount := 0;
    // Progression jusqu'a X4 (deja home).
    FB(Enable := TRUE, PowerContactorEngaged := TRUE, Mode := E_Mode.SEMI_AUTO,
       DeadmanArmed := TRUE, JoystickDeflected := TRUE, JoystickPush := TRUE, M1_SpeedValid := TRUE, M2_SpeedValid := TRUE, M1_ContactorsReleased := TRUE, M2_ContactorsReleased := TRUE, M1_BrakeApplied := TRUE, M2_BrakeApplied := TRUE, M1_SpeedStepApplied := 4, M2_SpeedStepApplied := 4, HeartbeatIhmOk := TRUE, StartCycle := TRUE,
       SelTarget := 3, LimitLegalDepthM := -10.5, CableLimitM1AscentM := 7.0, DiveStartMinM := 4.0,
       SpeedMismatchThresholdMps := 0.0, SpeedMismatchTimeout := T#0ms,
       HomedM1 := TRUE, HomedM2 := TRUE, InitPositionOk := TRUE, WinchesAtTopWindow := TRUE,
       M1_CablePosM := 7.0, M2_CablePosM := 7.0, Translation_At_P1 := TRUE, Translation_Done := TRUE,
       Benne_Done := FALSE, Benne_IsOpen := FALSE, Benne_IsClosed := TRUE, Benne_IsRoughlyClosed := TRUE,
       SampleCount := SampleCount);
    FB(Enable := TRUE, PowerContactorEngaged := TRUE, Mode := E_Mode.SEMI_AUTO,
       DeadmanArmed := TRUE, JoystickDeflected := TRUE, JoystickPush := TRUE, M1_SpeedValid := TRUE, M2_SpeedValid := TRUE, M1_ContactorsReleased := TRUE, M2_ContactorsReleased := TRUE, M1_BrakeApplied := TRUE, M2_BrakeApplied := TRUE, M1_SpeedStepApplied := 4, M2_SpeedStepApplied := 4, HeartbeatIhmOk := TRUE, StartCycle := FALSE,
       SelTarget := 3, LimitLegalDepthM := -10.5, CableLimitM1AscentM := 7.0, DiveStartMinM := 4.0,
       SpeedMismatchThresholdMps := 0.0, SpeedMismatchTimeout := T#0ms,
       HomedM1 := TRUE, HomedM2 := TRUE, InitPositionOk := TRUE, WinchesAtTopWindow := TRUE,
       M1_CablePosM := 7.0, M2_CablePosM := 7.0, Translation_At_P1 := TRUE, Translation_Done := TRUE,
       Benne_Done := FALSE, Benne_IsOpen := FALSE, Benne_IsClosed := TRUE, Benne_IsRoughlyClosed := TRUE,
       SampleCount := SampleCount);
    FB(Enable := TRUE, PowerContactorEngaged := TRUE, Mode := E_Mode.SEMI_AUTO,
       DeadmanArmed := TRUE, JoystickDeflected := TRUE, JoystickPush := TRUE, M1_SpeedValid := TRUE, M2_SpeedValid := TRUE, M1_ContactorsReleased := TRUE, M2_ContactorsReleased := TRUE, M1_BrakeApplied := TRUE, M2_BrakeApplied := TRUE, M1_SpeedStepApplied := 4, M2_SpeedStepApplied := 4, HeartbeatIhmOk := TRUE, StartCycle := FALSE,
       SelTarget := 3, LimitLegalDepthM := -10.5, CableLimitM1AscentM := 7.0, DiveStartMinM := 4.0,
       SpeedMismatchThresholdMps := 0.0, SpeedMismatchTimeout := T#0ms,
       HomedM1 := TRUE, HomedM2 := TRUE, InitPositionOk := TRUE, WinchesAtTopWindow := TRUE,
       M1_CablePosM := 7.0, M2_CablePosM := 7.0, Translation_At_P1 := TRUE, Translation_Done := TRUE,
       Benne_Done := TRUE, Benne_IsOpen := TRUE, Benne_IsClosed := FALSE, Benne_IsRoughlyClosed := FALSE,
       SampleCount := SampleCount);
    FB(Enable := TRUE, PowerContactorEngaged := TRUE, Mode := E_Mode.SEMI_AUTO,
       DeadmanArmed := TRUE, JoystickDeflected := TRUE, JoystickPush := TRUE, M1_SpeedValid := TRUE, M2_SpeedValid := TRUE, M1_ContactorsReleased := TRUE, M2_ContactorsReleased := TRUE, M1_BrakeApplied := TRUE, M2_BrakeApplied := TRUE, M1_SpeedStepApplied := 4, M2_SpeedStepApplied := 4, HeartbeatIhmOk := TRUE, StartCycle := FALSE,
       SelTarget := 3, LimitLegalDepthM := -10.5, CableLimitM1AscentM := 7.0, DiveStartMinM := 4.0,
       SpeedMismatchThresholdMps := 0.0, SpeedMismatchTimeout := T#0ms,
       HomedM1 := TRUE, HomedM2 := TRUE, InitPositionOk := TRUE, WinchesAtTopWindow := TRUE,
       M1_CablePosM := 5.0, M2_CablePosM := 5.0, Translation_At_P1 := TRUE, Translation_Done := TRUE,
       Benne_Done := TRUE, Benne_IsOpen := TRUE, Benne_IsClosed := FALSE, Benne_IsRoughlyClosed := FALSE,
       SampleCount := SampleCount);
    FB(Enable := TRUE, PowerContactorEngaged := TRUE, Mode := E_Mode.SEMI_AUTO,
       DeadmanArmed := TRUE, JoystickDeflected := TRUE, JoystickPush := TRUE, M1_SpeedValid := TRUE, M2_SpeedValid := TRUE, M1_ContactorsReleased := TRUE, M2_ContactorsReleased := TRUE, M1_BrakeApplied := TRUE, M2_BrakeApplied := TRUE, M1_SpeedStepApplied := 4, M2_SpeedStepApplied := 4, HeartbeatIhmOk := TRUE, StartCycle := FALSE,
       SelTarget := 3, LimitLegalDepthM := -10.5, CableLimitM1AscentM := 7.0, DiveStartMinM := 4.0,
       SpeedMismatchThresholdMps := 0.0, SpeedMismatchTimeout := T#0ms,
       HomedM1 := TRUE, HomedM2 := TRUE, InitPositionOk := TRUE, WinchesAtTopWindow := TRUE,
       M1_CablePosM := 5.0, M2_CablePosM := 5.0, Translation_At_P1 := TRUE, Translation_Done := TRUE,
       Benne_Done := TRUE, Benne_IsOpen := TRUE, Benne_IsClosed := FALSE, Benne_IsRoughlyClosed := FALSE,
       SampleCount := SampleCount);
    ADVANCE_TIME(300000000);
    FB(SampleCount := SampleCount);
    FB(SampleCount := SampleCount);
    ASSERT_TRUE(FB.CycleStep = E_AutoCycleStep.AX4_DESCEND_DIVING, 'Etabli en X4');
    // 40 s en X4 (< 60 s) -> pas de timeout.
    ADVANCE_TIME(40000000000);
    FB(Enable := TRUE, PowerContactorEngaged := TRUE, Mode := E_Mode.SEMI_AUTO,
       DeadmanArmed := TRUE, JoystickDeflected := TRUE, JoystickPush := TRUE, M1_SpeedValid := TRUE, M2_SpeedValid := TRUE, M1_ContactorsReleased := TRUE, M2_ContactorsReleased := TRUE, M1_BrakeApplied := TRUE, M2_BrakeApplied := TRUE, M1_SpeedStepApplied := 4, M2_SpeedStepApplied := 4, HeartbeatIhmOk := TRUE, StartCycle := FALSE,
       SelTarget := 3, LimitLegalDepthM := -10.5, CableLimitM1AscentM := 7.0, DiveStartMinM := 4.0,
       SpeedMismatchThresholdMps := 0.0, SpeedMismatchTimeout := T#0ms,
       HomedM1 := TRUE, HomedM2 := TRUE, InitPositionOk := TRUE, WinchesAtTopWindow := TRUE,
       M1_CablePosM := 5.0, M2_CablePosM := 5.0, Translation_At_P1 := TRUE, Translation_Done := TRUE,
       Benne_Done := TRUE, Benne_IsOpen := TRUE, Benne_IsClosed := FALSE, Benne_IsRoughlyClosed := FALSE,
       SampleCount := SampleCount);
    ASSERT_FALSE(FB.Fault.Error, 'X4 40 s : pas de timeout (< 60 s)');
    ASSERT_TRUE(FB.CycleStep = E_AutoCycleStep.AX4_DESCEND_DIVING, 'Toujours X4');
    // Contact fond -> X5. Nouvelle etape -> StepMaxTimer REARMEE (pas de cumul des 40 s de X4).
    FB(Enable := TRUE, PowerContactorEngaged := TRUE, Mode := E_Mode.SEMI_AUTO,
       DeadmanArmed := TRUE, JoystickDeflected := TRUE, JoystickPush := TRUE, M1_SpeedValid := TRUE, M2_SpeedValid := TRUE, M1_ContactorsReleased := TRUE, M2_ContactorsReleased := TRUE, M1_BrakeApplied := TRUE, M2_BrakeApplied := TRUE, M1_SpeedStepApplied := 4, M2_SpeedStepApplied := 4, HeartbeatIhmOk := TRUE, StartCycle := FALSE,
       SelTarget := 3, LimitLegalDepthM := -10.5, CableLimitM1AscentM := 7.0, DiveStartMinM := 4.0,
       SpeedMismatchThresholdMps := 0.0, SpeedMismatchTimeout := T#0ms,
       HomedM1 := TRUE, HomedM2 := TRUE, InitPositionOk := TRUE, WinchesAtTopWindow := TRUE,
       M1_CablePosM := 5.0, M2_CablePosM := 5.0, Translation_At_P1 := TRUE, Translation_Done := TRUE,
       Benne_Done := TRUE, Benne_IsOpen := TRUE, Benne_IsClosed := FALSE, Benne_IsRoughlyClosed := FALSE,
       SampleCount := SampleCount);
    // 1 scan de stabilisation en X5 pour armer StepMaxTimer sur la nouvelle etape.
    FB(Enable := TRUE, PowerContactorEngaged := TRUE, Mode := E_Mode.SEMI_AUTO,
       DeadmanArmed := TRUE, JoystickDeflected := TRUE, JoystickPush := TRUE, M1_SpeedValid := TRUE, M2_SpeedValid := TRUE, M1_ContactorsReleased := TRUE, M2_ContactorsReleased := TRUE, M1_BrakeApplied := TRUE, M2_BrakeApplied := TRUE, M1_SpeedStepApplied := 4, M2_SpeedStepApplied := 4, HeartbeatIhmOk := TRUE, StartCycle := FALSE,
       SelTarget := 3, LimitLegalDepthM := -10.5, CableLimitM1AscentM := 7.0, DiveStartMinM := 4.0,
       SpeedMismatchThresholdMps := 0.0, SpeedMismatchTimeout := T#0ms,
       HomedM1 := TRUE, HomedM2 := TRUE, InitPositionOk := TRUE, WinchesAtTopWindow := TRUE,
       M1_CablePosM := 5.0, M2_CablePosM := 5.0, Translation_At_P1 := TRUE, Translation_Done := TRUE,
       Benne_Done := TRUE, Benne_IsOpen := TRUE, Benne_IsClosed := FALSE, Benne_IsRoughlyClosed := FALSE,
       SampleCount := SampleCount);
    ASSERT_TRUE(FB.CycleStep = E_AutoCycleStep.AX4_DESCEND_DIVING, 'Etabli en AX4 (plongee)');
    // 40 s en X5 (< 60 s) -> total cycle 80 s mais aucune etape > 60 s -> PAS de AX_STAB.
    ADVANCE_TIME(40000000000);
    FB(Enable := TRUE, PowerContactorEngaged := TRUE, Mode := E_Mode.SEMI_AUTO,
       DeadmanArmed := TRUE, JoystickDeflected := TRUE, JoystickPush := TRUE, M1_SpeedValid := TRUE, M2_SpeedValid := TRUE, M1_ContactorsReleased := TRUE, M2_ContactorsReleased := TRUE, M1_BrakeApplied := TRUE, M2_BrakeApplied := TRUE, M1_SpeedStepApplied := 4, M2_SpeedStepApplied := 4, HeartbeatIhmOk := TRUE, StartCycle := FALSE,
       SelTarget := 3, LimitLegalDepthM := -10.5, CableLimitM1AscentM := 7.0, DiveStartMinM := 4.0,
       SpeedMismatchThresholdMps := 0.0, SpeedMismatchTimeout := T#0ms,
       HomedM1 := TRUE, HomedM2 := TRUE, InitPositionOk := TRUE, WinchesAtTopWindow := TRUE,
       M1_CablePosM := 5.0, M2_CablePosM := 5.0, Translation_At_P1 := TRUE, Translation_Done := TRUE,
       Benne_Done := TRUE, Benne_IsOpen := TRUE, Benne_IsClosed := FALSE, Benne_IsRoughlyClosed := FALSE,
       SampleCount := SampleCount);
    ASSERT_FALSE(FB.Fault.Error, 'X5 40 s : pas de timeout - StepMaxTimer non cumulatif sur le cycle');
    ASSERT_TRUE(FB.CycleStep = E_AutoCycleStep.AX4_DESCEND_DIVING, 'Toujours AX4, pas de AX_STAB (StepMaxTimer non cumulatif)');
END_TEST

TEST 'TC-P04-026 : AX4 ne contient aucun seuil synchro local - PRG04 reste source unique'
    SampleCount := 0;
    FB(Enable := TRUE, PowerContactorEngaged := TRUE, Mode := E_Mode.SEMI_AUTO,
       DeadmanArmed := TRUE, JoystickDeflected := TRUE, JoystickPush := TRUE, M1_SpeedValid := TRUE, M2_SpeedValid := TRUE, M1_ContactorsReleased := TRUE, M2_ContactorsReleased := TRUE, M1_BrakeApplied := TRUE, M2_BrakeApplied := TRUE, M1_SpeedStepApplied := 4, M2_SpeedStepApplied := 4, HeartbeatIhmOk := TRUE, StartCycle := TRUE,
       SelTarget := 3, LimitLegalDepthM := -10.5, CableLimitM1AscentM := 7.0,
       SpeedMismatchThresholdMps := 0.0, SpeedMismatchTimeout := T#0ms,
       HomedM1 := TRUE, HomedM2 := TRUE, InitPositionOk := TRUE, WinchesAtTopWindow := TRUE,
       M1_CablePosM := 7.0, M2_CablePosM := 7.0, Translation_At_P1 := TRUE, Translation_Done := TRUE,
       Benne_Done := FALSE, Benne_IsOpen := FALSE, Benne_IsClosed := TRUE, Benne_IsRoughlyClosed := TRUE,
       SampleCount := SampleCount);
    FB(Enable := TRUE, PowerContactorEngaged := TRUE, Mode := E_Mode.SEMI_AUTO,
       DeadmanArmed := TRUE, JoystickDeflected := TRUE, JoystickPush := TRUE, M1_SpeedValid := TRUE, M2_SpeedValid := TRUE, M1_ContactorsReleased := TRUE, M2_ContactorsReleased := TRUE, M1_BrakeApplied := TRUE, M2_BrakeApplied := TRUE, M1_SpeedStepApplied := 4, M2_SpeedStepApplied := 4, HeartbeatIhmOk := TRUE, StartCycle := FALSE,
       SelTarget := 3, LimitLegalDepthM := -10.5, CableLimitM1AscentM := 7.0,
       SpeedMismatchThresholdMps := 0.0, SpeedMismatchTimeout := T#0ms,
       HomedM1 := TRUE, HomedM2 := TRUE, InitPositionOk := TRUE, WinchesAtTopWindow := TRUE,
       M1_CablePosM := 7.0, M2_CablePosM := 7.0, Translation_At_P1 := TRUE, Translation_Done := TRUE,
       Benne_Done := FALSE, Benne_IsOpen := FALSE, Benne_IsClosed := TRUE, Benne_IsRoughlyClosed := TRUE,
       SampleCount := SampleCount);
    FB(Enable := TRUE, PowerContactorEngaged := TRUE, Mode := E_Mode.SEMI_AUTO,
       DeadmanArmed := TRUE, JoystickDeflected := TRUE, JoystickPush := TRUE, M1_SpeedValid := TRUE, M2_SpeedValid := TRUE, M1_ContactorsReleased := TRUE, M2_ContactorsReleased := TRUE, M1_BrakeApplied := TRUE, M2_BrakeApplied := TRUE, M1_SpeedStepApplied := 4, M2_SpeedStepApplied := 4, HeartbeatIhmOk := TRUE, StartCycle := FALSE,
       SelTarget := 3, LimitLegalDepthM := -10.5, CableLimitM1AscentM := 7.0,
       SpeedMismatchThresholdMps := 0.0, SpeedMismatchTimeout := T#0ms,
       HomedM1 := TRUE, HomedM2 := TRUE, InitPositionOk := TRUE, WinchesAtTopWindow := TRUE,
       M1_CablePosM := 7.0, M2_CablePosM := 7.0, Translation_At_P1 := TRUE, Translation_Done := TRUE,
       Benne_Done := TRUE, Benne_IsOpen := TRUE, Benne_IsClosed := FALSE, Benne_IsRoughlyClosed := FALSE,
       SampleCount := SampleCount);
    FB(Enable := TRUE, PowerContactorEngaged := TRUE, Mode := E_Mode.SEMI_AUTO,
       DeadmanArmed := TRUE, JoystickDeflected := TRUE, JoystickPush := TRUE, M1_SpeedValid := TRUE, M2_SpeedValid := TRUE, M1_ContactorsReleased := TRUE, M2_ContactorsReleased := TRUE, M1_BrakeApplied := TRUE, M2_BrakeApplied := TRUE, M1_SpeedStepApplied := 4, M2_SpeedStepApplied := 4, HeartbeatIhmOk := TRUE, StartCycle := FALSE,
       SelTarget := 3, LimitLegalDepthM := -10.5, CableLimitM1AscentM := 7.0,
       SpeedMismatchThresholdMps := 0.0, SpeedMismatchTimeout := T#0ms,
       HomedM1 := TRUE, HomedM2 := TRUE, InitPositionOk := TRUE, WinchesAtTopWindow := TRUE,
       M1_CablePosM := 5.0, M2_CablePosM := 5.0, Translation_At_P1 := TRUE, Translation_Done := TRUE,
       Benne_Done := TRUE, Benne_IsOpen := TRUE, Benne_IsClosed := FALSE, Benne_IsRoughlyClosed := FALSE,
       SampleCount := SampleCount);
    FB(Enable := TRUE, PowerContactorEngaged := TRUE, Mode := E_Mode.SEMI_AUTO,
       DeadmanArmed := TRUE, JoystickDeflected := TRUE, JoystickPush := TRUE, M1_SpeedValid := TRUE, M2_SpeedValid := TRUE, M1_ContactorsReleased := TRUE, M2_ContactorsReleased := TRUE, M1_BrakeApplied := TRUE, M2_BrakeApplied := TRUE, M1_SpeedStepApplied := 4, M2_SpeedStepApplied := 4, HeartbeatIhmOk := TRUE, StartCycle := FALSE,
       SelTarget := 3, LimitLegalDepthM := -10.5, CableLimitM1AscentM := 7.0,
       SpeedMismatchThresholdMps := 0.0, SpeedMismatchTimeout := T#0ms,
       HomedM1 := TRUE, HomedM2 := TRUE, InitPositionOk := TRUE, WinchesAtTopWindow := TRUE,
       M1_CablePosM := 5.0, M2_CablePosM := 5.0, Translation_At_P1 := TRUE, Translation_Done := TRUE,
       Benne_Done := TRUE, Benne_IsOpen := TRUE, Benne_IsClosed := FALSE, Benne_IsRoughlyClosed := FALSE,
       SampleCount := SampleCount);
    ADVANCE_TIME(300000000);
    FB(SampleCount := SampleCount);
    FB(SampleCount := SampleCount);
    ASSERT_TRUE(FB.CycleStep = E_AutoCycleStep.AX4_DESCEND_DIVING, 'Etabli en X4');
    // AX4..AX7 ne lisent aucun seuil de delta. PRG04 convertit ses causes critiques
    // (synchro confirmee, contacteurs ou Meca E) en WinchSyncError avant le cycle.
    FB(Enable := TRUE, PowerContactorEngaged := TRUE, Mode := E_Mode.SEMI_AUTO,
       DeadmanArmed := TRUE, JoystickDeflected := TRUE, JoystickPush := TRUE, M1_SpeedValid := TRUE, M2_SpeedValid := TRUE, M1_ContactorsReleased := TRUE, M2_ContactorsReleased := TRUE, M1_BrakeApplied := TRUE, M2_BrakeApplied := TRUE, M1_SpeedStepApplied := 4, M2_SpeedStepApplied := 4, HeartbeatIhmOk := TRUE, StartCycle := FALSE,
       SelTarget := 3, LimitLegalDepthM := -10.5, CableLimitM1AscentM := 7.0,
       SpeedMismatchThresholdMps := 0.0, SpeedMismatchTimeout := T#0ms,
       HomedM1 := TRUE, HomedM2 := TRUE, InitPositionOk := TRUE, WinchesAtTopWindow := TRUE,
       M1_CablePosM := 5.0, M2_CablePosM := 5.0,
       WinchSyncError := FALSE, WinchSyncDeltaM := 0.0,
       Translation_At_P1 := TRUE, Translation_Done := TRUE,
       Benne_Done := TRUE, Benne_IsOpen := TRUE, Benne_IsClosed := FALSE, Benne_IsRoughlyClosed := FALSE,
       SampleCount := SampleCount);
    ASSERT_TRUE(FB.CycleStep = E_AutoCycleStep.AX4_DESCEND_DIVING, 'AX4 reste pilote uniquement par WinchSyncError PRG04');
    ASSERT_FALSE(FB.Fault.Error, 'Aucun seuil synchro local cycle');
END_TEST

TEST 'TC-P04-022 : Abort+Start avec Fault.Latched actif -> cycle reste en X0 (pas de redemarrage) (T192-A S1)'
    SampleCount := 0;
    // Scan 1 : Demarrage (front StartCycle) -> X0 vers X1
    FB(Enable := TRUE, PowerContactorEngaged := TRUE, Mode := E_Mode.SEMI_AUTO,
       DeadmanArmed := TRUE, JoystickDeflected := TRUE, JoystickPush := TRUE, M1_SpeedValid := TRUE, M2_SpeedValid := TRUE, M1_ContactorsReleased := TRUE, M2_ContactorsReleased := TRUE, M1_BrakeApplied := TRUE, M2_BrakeApplied := TRUE, M1_SpeedStepApplied := 4, M2_SpeedStepApplied := 4, HeartbeatIhmOk := TRUE,
       StartCycle := TRUE, AbortCycle := FALSE, WinchSyncError := FALSE, Reset := FALSE,
       HomedM1 := FALSE, HomedM2 := FALSE, HomingRequest := FALSE,
       M1_CablePosM := -10.0, M2_CablePosM := -10.0, M1_MeasuredSpeedMps := 0.0, M2_MeasuredSpeedMps := 0.0,
       SpeedMismatchThresholdMps := 0.0, SpeedMismatchTimeout := T#0ms,
WinchSyncDeltaM := 0.0,
       Translation_At_P1 := FALSE, Translation_At_Tremie := FALSE, Translation_At_Maintenance := FALSE,
       Translation_Busy := FALSE, Translation_Done := FALSE,
       Benne_Busy := FALSE, Benne_Done := FALSE, Benne_IsOpen := FALSE, Benne_IsClosed := FALSE, Benne_IsRoughlyClosed := FALSE,
       SampleCount := SampleCount);
    // Scan 2 : StartCycle relache -> etablissement AX1_INIT
    FB(Enable := TRUE, PowerContactorEngaged := TRUE, Mode := E_Mode.SEMI_AUTO,
       DeadmanArmed := TRUE, JoystickDeflected := TRUE, JoystickPush := TRUE, M1_SpeedValid := TRUE, M2_SpeedValid := TRUE, M1_ContactorsReleased := TRUE, M2_ContactorsReleased := TRUE, M1_BrakeApplied := TRUE, M2_BrakeApplied := TRUE, M1_SpeedStepApplied := 4, M2_SpeedStepApplied := 4, HeartbeatIhmOk := TRUE,
       StartCycle := FALSE, AbortCycle := FALSE, WinchSyncError := FALSE, Reset := FALSE,
       HomedM1 := FALSE, HomedM2 := FALSE, HomingRequest := FALSE,
       M1_CablePosM := -10.0, M2_CablePosM := -10.0, M1_MeasuredSpeedMps := 0.0, M2_MeasuredSpeedMps := 0.0,
       SpeedMismatchThresholdMps := 0.0, SpeedMismatchTimeout := T#0ms,
WinchSyncDeltaM := 0.0,
       Translation_At_P1 := FALSE, Translation_At_Tremie := FALSE, Translation_At_Maintenance := FALSE,
       Translation_Busy := FALSE, Translation_Done := FALSE,
       Benne_Busy := FALSE, Benne_Done := FALSE, Benne_IsOpen := FALSE, Benne_IsClosed := FALSE, Benne_IsRoughlyClosed := FALSE,
       SampleCount := SampleCount);
    ASSERT_TRUE(FB.CycleStep = E_AutoCycleStep.AX1_INIT, 'Etablissement a AX1_INIT');
    // Scan 3 : Injection defaut synchronisme -> AX_STAB + Fault.Latched=TRUE
    FB(Enable := TRUE, PowerContactorEngaged := TRUE, Mode := E_Mode.SEMI_AUTO,
       DeadmanArmed := TRUE, JoystickDeflected := TRUE, JoystickPush := TRUE, M1_SpeedValid := TRUE, M2_SpeedValid := TRUE, M1_ContactorsReleased := TRUE, M2_ContactorsReleased := TRUE, M1_BrakeApplied := TRUE, M2_BrakeApplied := TRUE, M1_SpeedStepApplied := 4, M2_SpeedStepApplied := 4, HeartbeatIhmOk := TRUE,
       StartCycle := FALSE, AbortCycle := FALSE, WinchSyncError := TRUE, Reset := FALSE,
       HomedM1 := FALSE, HomedM2 := FALSE, HomingRequest := FALSE,
       M1_CablePosM := -10.0, M2_CablePosM := -10.0, M1_MeasuredSpeedMps := 0.0, M2_MeasuredSpeedMps := 0.0,
       SpeedMismatchThresholdMps := 0.0, SpeedMismatchTimeout := T#0ms,
WinchSyncDeltaM := 0.0,
       Translation_At_P1 := FALSE, Translation_At_Tremie := FALSE, Translation_At_Maintenance := FALSE,
       Translation_Busy := FALSE, Translation_Done := FALSE,
       Benne_Busy := FALSE, Benne_Done := FALSE, Benne_IsOpen := FALSE, Benne_IsClosed := FALSE, Benne_IsRoughlyClosed := FALSE,
       SampleCount := SampleCount);
    ASSERT_TRUE(FB.CycleStep = E_AutoCycleStep.AX_STAB, 'Bascule en AX_STAB sur defaut');
    ASSERT_TRUE(FB.Fault.Latched, 'Defaut latche actif');
    // Scan 4 : Cause disparue (Error retombe) mais Latch persiste (pas de Reset)
    FB(Enable := TRUE, PowerContactorEngaged := TRUE, Mode := E_Mode.SEMI_AUTO,
       DeadmanArmed := TRUE, JoystickDeflected := TRUE, JoystickPush := TRUE, M1_SpeedValid := TRUE, M2_SpeedValid := TRUE, M1_ContactorsReleased := TRUE, M2_ContactorsReleased := TRUE, M1_BrakeApplied := TRUE, M2_BrakeApplied := TRUE, M1_SpeedStepApplied := 4, M2_SpeedStepApplied := 4, HeartbeatIhmOk := TRUE,
       StartCycle := FALSE, AbortCycle := FALSE, WinchSyncError := FALSE, Reset := FALSE,
       HomedM1 := FALSE, HomedM2 := FALSE, HomingRequest := FALSE,
       M1_CablePosM := -10.0, M2_CablePosM := -10.0, M1_MeasuredSpeedMps := 0.0, M2_MeasuredSpeedMps := 0.0,
       SpeedMismatchThresholdMps := 0.0, SpeedMismatchTimeout := T#0ms,
WinchSyncDeltaM := 0.0,
       Translation_At_P1 := FALSE, Translation_At_Tremie := FALSE, Translation_At_Maintenance := FALSE,
       Translation_Busy := FALSE, Translation_Done := FALSE,
       Benne_Busy := FALSE, Benne_Done := FALSE, Benne_IsOpen := FALSE, Benne_IsClosed := FALSE, Benne_IsRoughlyClosed := FALSE,
       SampleCount := SampleCount);
    ASSERT_TRUE(FB.Fault.Latched, 'Latch persiste sans Reset');
    // Scan 5 : AbortCycle -> retour X0 (mais Latch toujours actif)
    FB(Enable := TRUE, PowerContactorEngaged := TRUE, Mode := E_Mode.SEMI_AUTO,
       DeadmanArmed := TRUE, JoystickDeflected := TRUE, JoystickPush := TRUE, M1_SpeedValid := TRUE, M2_SpeedValid := TRUE, M1_ContactorsReleased := TRUE, M2_ContactorsReleased := TRUE, M1_BrakeApplied := TRUE, M2_BrakeApplied := TRUE, M1_SpeedStepApplied := 4, M2_SpeedStepApplied := 4, HeartbeatIhmOk := TRUE,
       StartCycle := FALSE, AbortCycle := TRUE, WinchSyncError := FALSE, Reset := FALSE,
       HomedM1 := FALSE, HomedM2 := FALSE, HomingRequest := FALSE,
       M1_CablePosM := -10.0, M2_CablePosM := -10.0, M1_MeasuredSpeedMps := 0.0, M2_MeasuredSpeedMps := 0.0,
       SpeedMismatchThresholdMps := 0.0, SpeedMismatchTimeout := T#0ms,
WinchSyncDeltaM := 0.0,
       Translation_At_P1 := FALSE, Translation_At_Tremie := FALSE, Translation_At_Maintenance := FALSE,
       Translation_Busy := FALSE, Translation_Done := FALSE,
       Benne_Busy := FALSE, Benne_Done := FALSE, Benne_IsOpen := FALSE, Benne_IsClosed := FALSE, Benne_IsRoughlyClosed := FALSE,
       SampleCount := SampleCount);
    ASSERT_TRUE(FB.CycleStep = E_AutoCycleStep.AX0_REPOS, 'Abort -> retour X0');
    // Scan 6 : StartCycle avec Fault.Latched actif -> RESTE EN X0 (gate NOT Fault.Latched)
    FB(Enable := TRUE, PowerContactorEngaged := TRUE, Mode := E_Mode.SEMI_AUTO,
       DeadmanArmed := TRUE, JoystickDeflected := TRUE, JoystickPush := TRUE, M1_SpeedValid := TRUE, M2_SpeedValid := TRUE, M1_ContactorsReleased := TRUE, M2_ContactorsReleased := TRUE, M1_BrakeApplied := TRUE, M2_BrakeApplied := TRUE, M1_SpeedStepApplied := 4, M2_SpeedStepApplied := 4, HeartbeatIhmOk := TRUE,
       StartCycle := TRUE, AbortCycle := FALSE, WinchSyncError := FALSE, Reset := FALSE,
       HomedM1 := FALSE, HomedM2 := FALSE, HomingRequest := FALSE,
       M1_CablePosM := -10.0, M2_CablePosM := -10.0, M1_MeasuredSpeedMps := 0.0, M2_MeasuredSpeedMps := 0.0,
       SpeedMismatchThresholdMps := 0.0, SpeedMismatchTimeout := T#0ms,
WinchSyncDeltaM := 0.0,
       Translation_At_P1 := FALSE, Translation_At_Tremie := FALSE, Translation_At_Maintenance := FALSE,
       Translation_Busy := FALSE, Translation_Done := FALSE,
       Benne_Busy := FALSE, Benne_Done := FALSE, Benne_IsOpen := FALSE, Benne_IsClosed := FALSE, Benne_IsRoughlyClosed := FALSE,
       SampleCount := SampleCount);
    ASSERT_TRUE(FB.CycleStep = E_AutoCycleStep.AX0_REPOS, 'Reste en X0 : Start bloque par Fault.Latched (S1)');
    // Scan 7 : StartCycle relache -> confirme X0, pas de redemarrage
    FB(Enable := TRUE, PowerContactorEngaged := TRUE, Mode := E_Mode.SEMI_AUTO,
       DeadmanArmed := TRUE, JoystickDeflected := TRUE, JoystickPush := TRUE, M1_SpeedValid := TRUE, M2_SpeedValid := TRUE, M1_ContactorsReleased := TRUE, M2_ContactorsReleased := TRUE, M1_BrakeApplied := TRUE, M2_BrakeApplied := TRUE, M1_SpeedStepApplied := 4, M2_SpeedStepApplied := 4, HeartbeatIhmOk := TRUE,
       StartCycle := FALSE, AbortCycle := FALSE, WinchSyncError := FALSE, Reset := FALSE,
       HomedM1 := FALSE, HomedM2 := FALSE, HomingRequest := FALSE,
       M1_CablePosM := -10.0, M2_CablePosM := -10.0, M1_MeasuredSpeedMps := 0.0, M2_MeasuredSpeedMps := 0.0,
       SpeedMismatchThresholdMps := 0.0, SpeedMismatchTimeout := T#0ms,
WinchSyncDeltaM := 0.0,
       Translation_At_P1 := FALSE, Translation_At_Tremie := FALSE, Translation_At_Maintenance := FALSE,
       Translation_Busy := FALSE, Translation_Done := FALSE,
       Benne_Busy := FALSE, Benne_Done := FALSE, Benne_IsOpen := FALSE, Benne_IsClosed := FALSE, Benne_IsRoughlyClosed := FALSE,
       SampleCount := SampleCount);
    ASSERT_TRUE(FB.CycleStep = E_AutoCycleStep.AX0_REPOS, 'Confirme X0 apres Start relache');
    ASSERT_FALSE(FB.Lifecycle.Busy, 'Pas de cycle en cours (Busy=FALSE)');
END_TEST
